(* IEC 61131-3 sources: daoli-st-library/DL_Base (part 15) *)

(* ---- FB_DL_RailPowerSequence.st ---- *)
(*
  ==================================================================
  组件名 Component  : FB_DL_RailPowerSequence
  分类   Category   : DL_Base
  前缀   Naming     : FB_DL_ ｜ b/n/u/f/t/e/st 类型前缀制（R265）
  复杂度 Complexity  : 中
  版本   Version    : 1.0.3
  功能   Purpose    : 多路供电轨按序上电/断电（延时可配、断电逆序、步进超时锁存）。
  来源   Source     : self-std（供电时序公开工程语义自研）
  平台   Platform   : 纯 IEC 61131-3（TON / R_TRIG / CASE），三平台通用
  分工声明 Split     : 与 FB_DL_LaserWeldPowerSeq（工艺专用属主）分工——后者绑定
                      激光焊接工艺流；本件为通用时序原子，不绑工艺、不判负载
                      特性（R216 双向互引）。
  作者   Author     : 道莅代码库 · PLC 编程专家（R61）
  归属 Ownership     : E_DL_RailPhase 属主为本文件（全库唯一定义，R264）；
                      引用件只引用不重声明。
  ------------------------------------------------------------------
  边界 Boundary     :
                      一 uRailCount = 0 或 > 8 判组态非法故障码，不进时序
                         （边界五；R239 显式分支，禁比较算子隐式分流）；
                      二 断电逆序强制：断电步序 = 上电步序倒序（结构写死）；
                      三 步进超时按「单轨」计时（v1.0.2 修 D2）：tonStep.IN 串入逐拍派生
                         的本轨待响应量 _bRailPending（eRampUp 取 NOT abRailFb[_nStep]、
                         eRampDn 取 abRailFb[_nStep]），本轨一响应即自动复位，不再整段
                         连续计时；锁存独立码 + 解除式可达自证：故障相由复位沿迁回空闲
                         并清锁存（bReset 输入引脚恒可达，R152 自证）；
                      三A 上电推进判据「沿 OR 电平」双路（v1.0.3 修 R62-D4 中）：eRampUp
                         推进条件 = rtFb.Q（反馈上升沿）OR abRailFb[_nStep]（电平已就位
                         直过）——「反馈预闭合」处置口径：若轨在上一步计时期间或起步拍
                         前反馈电平已提前闭合（边沿被上一步消费 / 起步拍无沿），单轨超时
                         门控（_bRailPending = FALSE）与推进判据（仅沿）同源失效会静默
                         挂死；电平直过支路消除该挂死路径。断电相完成判据本为电平式
                         （NOT abRailFb[_nStep]），无此问题；
                      七 空轨断电早退（v1.0.2 修 D1）：_nCnt = 0 时收到断电沿不迁移、
                         不置 bDone、仅发信息级 0655，防伪造「完成单拍」；原负下标
                         钳位语句保留为二重防御，不再是唯一防线；
                      四 状态机 ENUM + CASE，ELSE 拦非法态；TON/R_TRIG 段 0
                         无条件刷新（禁入分支，R7）；TON IN 串故障锁存门控
                         （FB50-1）；
                      五 使能失电语义为「弃用本轮时序」（回空闲，不锁存不出
                         单拍）——R191 声明行；
                      六 无全局、无外部变量、无物理地址。
  错误码   Codes    :
    16#0001_0642【故障级】供电轨数组态非法（=0 或 >8），锁存至复位沿
    16#0001_0643【故障级】步进反馈超时（tStepTimeout 内未见该轨反馈），锁存至复位沿
    16#0001_0655【信息级】空轨断电请求已忽略（_nCnt 为 0 时无可断轨，不迁移不置 bDone）
  验收   Acceptance :
    算法已证（脚本）：未跑 ｜ 编译器已证（三平台）：未跑
    V1 3 轨、反馈逐轨到位 → uOnCount=3、bDone 单拍
    V2 第 2 轨反馈不至 → 码 0643、eFault、锁存待复位
    V3 uRailCount=0 → 码 0642、不进时序
    V4 空轨断电（abRailFb 全 FALSE、bOffCmd 上升沿）→ bDone 全拍 FALSE、
       eState 保持 eIdle、eErr=0655（v1.0.2 回归向量）
    V5 3 轨、每轨反馈延时 0.8×tStepTimeout → 全序列成功、无 0643；
       单轨延时 1.2× → 该轨锁 0643（v1.0.2 单轨超时回归向量）
    V6 轨 2 反馈预闭合（在轨 1 计时期间电平提前拉高，无沿）→ 轨 2 仍被推进、
       不锁 0643（v1.0.3 沿 OR 电平双路回归向量）
  修订记录 Revision  :
    2026-11-21  v1.0.0  R61 首版（批 3 · 序号 9）
    2026-11-21  v1.0.1  R61 终审 D1 就地修（安全侧）：空轨断电起步 _nStep<0 钳位、堵 abRailFb[-1] 越界读（R333 安全侧例外，正常路径行为零变更）
    2026-11-21  v1.0.2  R62-D1/D2 返修：①eIdle/eStable 的 rtOff 分支加 _nCnt=0 空轨早退（不迁移、不置 bDone、仅信息码 0655），原钳位降为二重防御；②新增 _bRailPending 串入 tonStep.IN 实现单轨超时；③段 0 rtFb 刷新条件扩到 eRampUp 或 eRampDn
    2026-11-21  v1.0.3  R63 返修 R4（R62-D4 中）：eRampUp 推进判据改「沿 OR 电平」双路（rtFb.Q OR abRailFb[_nStep]），反馈预闭合轨电平直过，消除单轨超时门控与推进判据同源静默挂死；头注释补「反馈预闭合」处置口径与向量 V6
  ==================================================================
*)
TYPE E_DL_RailPhase :
(
    eIdle    := 0,  // 空闲：等上电/断电命令沿 / idle, waiting for the power command edges
    eRampUp  := 10, // 上电步进：正向逐轨 / the power up stepping forward rail by rail
    eStable  := 20, // 稳定：全轨已上 / stable, all rails powered
    eRampDn  := 30  // 断电步进：逆向逐轨（边界二）/ the power down stepping in the reverse order
);
END_TYPE

FUNCTION_BLOCK FB_DL_RailPowerSequence
VAR_INPUT
    bOnCmd       : BOOL := FALSE; // 上电命令电平，上升沿发起正向时序 / the power on command level
    bOffCmd      : BOOL := FALSE; // 断电命令电平，上升沿发起逆向时序 / the power off command level
    bReset       : BOOL := FALSE; // 故障复位电平，上升沿清锁存回空闲 / the fault reset level
    uRailCount   : UDINT := 3;    // 供电轨数 [路]，合法域 1..8 / the rail count, legal from one to eight
    tStepTimeout : TIME := T#5S;  // 单轨步进超时 [毫秒] / the per rail step timeout
END_VAR
VAR_IN_OUT
    abRailFb  : ARRAY[0..7] OF BOOL; // 各轨反馈电平 [路反馈]，只读 / the rail feedback levels, read only
    atOnDelay : ARRAY[0..7] OF TIME; // 各轨上电前延时 [毫秒]，可配 / the per rail pre power delay, configurable
END_VAR
VAR_OUTPUT
    uOnCnt  : UDINT := 0;              // 已上电轨数 [路] / the powered rail count
    bDone   : BOOL := FALSE;           // 本轮时序完成单拍脉冲 [-] / the round done one shot pulse
    eState  : E_DL_RailPhase;          // 主状态机当前态 [状态] / the current state
    bError  : BOOL := FALSE;           // 故障锁存位（与锁存同源，R191）/ the fault bit from the latch
    eErr    : UDINT := 16#0000_0000;   // 错误码，0 = 正常 / the error code, zero is ok
END_VAR
VAR
    _bInit   : BOOL := FALSE;                          // 首拍初始化标志（R310）/ the first scan flag
    _eState  : E_DL_RailPhase := E_DL_RailPhase.eIdle; // 内部状态寄存器 / the internal state register
    _bDone   : BOOL := FALSE;                          // 完成单拍内部位，段 1 预清段 5 映射 / the internal done bit
    _bFault  : BOOL := FALSE;                          // 故障锁存副本（仅复位沿清除）/ the fault latch copy
    _nStep   : DINT  := 0;                             // 当前步进轨索引 [下标] / the current step rail index
    _nCnt    : UDINT := 0;                             // 已完成轨数副本 [路] / the completed rail count copy
    _nUse    : DINT  := 0;                             // 钳位后的轨数 [路] / the clamped rail count
    _bCfgBad : BOOL  := FALSE;                         // 组态非法标记（逐拍重算）/ the configuration fault flag
    _bStepGo : BOOL  := FALSE;                         // 步进计时使能（驻留派生）[-] / the step timing enable derived from the dwell
    _bRailPending : BOOL := FALSE;                     // 本轨待响应量（逐拍派生：上电取未反馈、断电取仍反馈）[-] / the pending rail of this step, derived every scan
    _bEmptyOff : BOOL := FALSE;                        // 空轨断电早退标记（逐拍重算，信息级 0655）/ the empty bank off request flag, recomputed every scan
    rtOn     : R_TRIG;  // 上电命令沿实例，段 0 无条件刷新 / the on command edge instance
    rtOff    : R_TRIG;  // 断电命令沿实例，段 0 无条件刷新 / the off command edge instance
    rtReset  : R_TRIG;  // 复位沿实例，段 0 无条件刷新 / the reset edge instance
    rtFb     : R_TRIG;  // 步进轨反馈沿实例，段 0 无条件刷新 / the step rail feedback edge instance
    tonStep  : TON;     // 步进超时计时器，段 0 无条件刷新 / the step timeout timer
END_VAR
VAR CONSTANT
    DL_RPS_RMAX : DINT := 8; // 供电轨容量上界 [路]，与数组容量一致 / the rail capacity aligned with the array
END_VAR

// 段 0｜定时器与沿检测无条件周期刷新（禁入分支，R7；TON IN 串故障锁存门控，FB50-1）/ segment 0, the unconditional refresh
rtOn(CLK := bOnCmd); // 上电沿 / the on edge
rtOff(CLK := bOffCmd); // 断电沿 / the off edge
rtReset(CLK := bReset); // 复位沿 / the reset edge
IF (_eState = E_DL_RailPhase.eRampUp) OR (_eState = E_DL_RailPhase.eRampDn) THEN // 两相步进相均刷当前轨反馈（v1.0.2 扩相，防断电相恒刷 0 号轨）/ both stepping phases watch the current rail
    rtFb(CLK := abRailFb[_nStep]); // 当前步进轨反馈沿 / the current step rail feedback edge
ELSE // 非步进相：非步进相固定刷新 0 号轨（保持无条件调用形态）/ the other phases refresh on the rail zero slot
    rtFb(CLK := abRailFb[0]); // 固定下标刷新 / the fixed index refresh
END_IF
_bStepGo := (_eState = E_DL_RailPhase.eRampUp) OR (_eState = E_DL_RailPhase.eRampDn); // 步进相驻留派生 / the dwell derived enable
// 单轨待响应量：只由「本相 + 本轨反馈」派生，本轨一响应即落 FALSE 使 TON 自动复位（v1.0.2 修 D2）/ the per rail pending, the timer resets by itself once this rail responds
IF _eState = E_DL_RailPhase.eRampUp THEN // 上电相：本轨尚未反馈即待响应 / the ramp up phase waits for the feedback to appear
    _bRailPending := NOT abRailFb[_nStep]; // 未反馈为待响应 / pending while the feedback is still absent
ELSIF _eState = E_DL_RailPhase.eRampDn THEN // 断电相：本轨仍反馈即待响应 / the ramp down phase waits for the feedback to vanish
    _bRailPending := abRailFb[_nStep]; // 仍反馈为待响应 / pending while the feedback is still present
ELSE // 其余相无单轨待响应语义 / no per rail pending outside the stepping phases
    _bRailPending := FALSE; // 非步进相清待响应 / clear the pending outside the stepping phases
END_IF
tonStep(IN := _bStepGo AND (NOT _bFault) AND _bRailPending, PT := tStepTimeout); // 单轨超时（串故障锁存门控 + 本轨待响应，FB50-1）/ the per rail timeout with the latch gate and the rail pending

// 段 1｜首拍初始化与单拍标志预清（FB32-1；R256）/ segment 1, the first scan init and the preset
IF NOT _bInit THEN // 首拍一拍 / the first scan
    _bInit := TRUE; // 置首拍标志 / raise the first scan flag
    _bFault := FALSE; // 故障锁存显式清零 / clear the fault latch explicitly
    _nStep := 0; // 步进索引显式清零 / clear the step index explicitly
    _nCnt := 0; // 完成轨数显式清零 / clear the completed count explicitly
    _eState := E_DL_RailPhase.eIdle; // 状态显式落空闲 / place the state to idle
END_IF
IF rtReset.Q THEN // 复位沿（作用域：清锁存 + 迁相位 + 清步进量，R311）/ the reset edge with the declared scope
    _bFault := FALSE; // 清故障锁存 / clear the fault latch
    _nStep := 0; // 清步进索引 / clear the step index
    _nCnt := 0; // 清完成轨数 / clear the completed count
    _eState := E_DL_RailPhase.eIdle; // 迁回空闲 / back to idle
END_IF
_bDone := FALSE; // 完成单拍预清零 / preset the done pulse false
_bCfgBad := FALSE; // 组态标记预清零 / preset the configuration flag false
_bEmptyOff := FALSE; // 空轨早退标记预清零（单拍信息位，段 5 映射 0655）/ preset the empty bank flag false

// 段 2｜组态域闸（轨数合法域 1..8，边界一）/ segment 2, the rail count gate
_nUse := UDINT_TO_DINT(uRailCount); // 轨数升位接管（超 DINT 域转负即被下界捕获）/ take the rail count widened, an overflow lands below the floor
IF (_nUse < 1) OR (_nUse > DL_RPS_RMAX) THEN // 轨数越域 / the rail count out of the domain
    _bCfgBad := TRUE; // 置组态非法标记 / raise the configuration flag
    _bFault := TRUE; // 锁存故障（0642，段 5 回放）/ latch the fault
END_IF
IF _nUse < 1 THEN // 下界钳位（防越界索引）/ the floor clamp for the index safety
    _nUse := 1; // 钳到一 / clamp to one
END_IF
IF _nUse > DL_RPS_RMAX THEN // 上界钳位 / the ceiling clamp
    _nUse := DL_RPS_RMAX; // 钳到容量 / clamp to the capacity
END_IF

// 段 3｜主状态机（ENUM + CASE，ELSE 拦非法态；安全相迁移带全量闸位复检，R274）/ segment 3, the main machine
CASE _eState OF
    E_DL_RailPhase.eIdle: // 空闲相 / the idle phase
        IF rtOn.Q AND (NOT _bFault) AND (NOT _bCfgBad) THEN // 上电沿 + 全量闸位复检（R274）/ the on edge with the full gate recheck
            _nStep := 0; // 从 0 号轨正向起步 / start forward from the rail zero
            _nCnt := 0; // 完成轨数归零 / reset the completed count
            _eState := E_DL_RailPhase.eRampUp; // 迁入上电步进相 / enter the ramp up phase
        ELSIF rtOff.Q AND (NOT _bFault) AND (NOT _bCfgBad) THEN // 断电沿 + 全量闸位复检 / the off edge with the recheck
            IF _nCnt = 0 THEN // 空轨早退（v1.0.2 修 D1）：无已上电轨则无从逆序断电 / the empty bank early exit, no powered rail to cut
                _bEmptyOff := TRUE; // 仅置信息级标记，不迁移、不置 bDone / raise the informational flag only, no migration and no done pulse
            ELSE // 有已上电轨：正常逆序起步 / a powered bank, start the reverse sequence
                _nStep := UDINT_TO_DINT(_nCnt) - 1; // 从已完成末轨逆向起步（断电逆序，边界二）/ start reverse from the last powered rail
                IF _nStep < 0 THEN // 二重防御：空轨已在上面早退，本钳位不再是唯一防线（R61-D1 保留）/ a second line of defence, no longer the only guard
                    _nStep := 0; // 钳到 0 号轨，防 abRailFb[-1] 越界读 / clamp to the rail zero against the negative index read
                END_IF
                _eState := E_DL_RailPhase.eRampDn; // 迁入断电步进相 / enter the ramp down phase
            END_IF
        END_IF
    E_DL_RailPhase.eRampUp: // 上电步进相 / the ramp up phase
        IF rtFb.Q OR abRailFb[_nStep] THEN // 推进判据「沿 OR 电平」双路（v1.0.3 修 R62-D4）：沿到或电平已预闭合均直过，防超时门控与推进判据同源静默挂死 / the advance criterion in the edge OR level dual path, a pre closed feedback passes by level so the timeout gate and the advance criterion cannot fail together in silence
            _nCnt := _nCnt + 1; // 完成轨数推进 / advance the completed count
            _nStep := _nStep + 1; // 步进索引推进 / advance the step index
            IF _nStep >= _nUse THEN // 全轨完成 / all rails done
                _bDone := TRUE; // 置完成单拍 / raise the done pulse
                _eState := E_DL_RailPhase.eStable; // 迁入稳定相 / enter the stable phase
            END_IF
        ELSIF tonStep.Q THEN // 步进超时（边界三）/ the step timeout
            _bFault := TRUE; // 锁存超时故障（0643）/ latch the timeout fault
        ELSIF _bFault THEN // 前置条件消失出口 / the prerequisite gone exit
            _eState := E_DL_RailPhase.eIdle; // 迁回空闲（锁存迁移由段 4 收口）/ back to idle
        END_IF
    E_DL_RailPhase.eStable: // 稳定相 / the stable phase
        IF rtOff.Q AND (NOT _bFault) THEN // 断电沿 + 闸位复检 / the off edge with the recheck
            IF _nCnt = 0 THEN // 空轨早退（与 eIdle 同口径，v1.0.2 修 D1）：异常态下 _nCnt 被清零亦不得伪造完成 / the same empty bank exit as the idle phase
                _bEmptyOff := TRUE; // 仅置信息级标记，不迁移、不置 bDone / raise the informational flag only
            ELSE // 有已上电轨：正常逆序起步 / a powered bank, start the reverse sequence
                _nStep := UDINT_TO_DINT(_nCnt) - 1; // 逆向起步（断电逆序）/ start reverse
                IF _nStep < 0 THEN // 二重防御（空轨已在上面早退）/ a second line of defence
                    _nStep := 0; // 钳到 0 号轨，防负下标越界读 / clamp to the rail zero against the negative index read
                END_IF
                _eState := E_DL_RailPhase.eRampDn; // 迁入断电步进相 / enter the ramp down phase
            END_IF
        ELSIF _bFault THEN // 前置条件消失 / the prerequisite gone
            _eState := E_DL_RailPhase.eIdle; // 迁回空闲 / back to idle
        END_IF
    E_DL_RailPhase.eRampDn: // 断电步进相（逆序，边界二）/ the ramp down phase in the reverse order
        IF NOT abRailFb[_nStep] THEN // 当前轨反馈已消失（断电完成判据）/ the current rail feedback gone
            IF _nCnt > 0 THEN // 无符号下溢闸（0 减 1 会回绕，先判再减）/ the underflow guard before the decrement
                _nCnt := _nCnt - 1; // 完成轨数回退 / step the completed count back
            END_IF
            _nStep := _nStep - 1; // 逆向推进 / step reverse
            IF _nStep < 0 THEN // 全轨断完 / all rails off
                _nCnt := 0; // 完成轨数清零 / clear the completed count
                _bDone := TRUE; // 置完成单拍 / raise the done pulse
                _eState := E_DL_RailPhase.eIdle; // 迁回空闲 / back to idle
            END_IF
        ELSIF tonStep.Q THEN // 步进超时 / the step timeout
            _bFault := TRUE; // 锁存超时故障 / latch the timeout fault
        ELSIF _bFault THEN // 前置条件消失 / the prerequisite gone
            _eState := E_DL_RailPhase.eIdle; // 迁回空闲 / back to idle
        END_IF
    ELSE // 非法枚举值拦截 / the illegal enumeration guard
        _eState := E_DL_RailPhase.eIdle; // 落回空闲 / force back to idle
        _bFault := TRUE; // 置故障锁存 / latch the fault
END_CASE

// 段 4｜故障锁存迁移闸（置于解除段之后防同拍抢迁，R258）/ segment 4, the latch to phase gate
IF _bFault AND (_eState <> E_DL_RailPhase.eIdle) THEN // 已锁存但不在空闲相（本件锁存即弃用本轮迁空闲）/ latched, the round is discarded to idle
    _eState := E_DL_RailPhase.eIdle; // 迁回空闲 / back to idle
END_IF

// 段 5｜统一出口（内部副本单点映射；故障码锁存回放，R187）/ segment 5, the unified outlet
uOnCnt := _nCnt; // 已上电轨数出口 / the powered count outlet
bDone := _bDone; // 完成单拍出口 / the done pulse outlet
eState := _eState; // 状态出口 / the state outlet
bError := _bFault; // 故障位出口（与锁存同源）/ the fault bit outlet
IF _bFault THEN // 故障锁存回放优先 / the latched fault replays first
    IF _bCfgBad THEN // 组态成因（独立码值，R190）/ the configuration cause
        eErr := 16#0001_0642; // 故障级：轨数组态非法 / fault grade, the illegal rail count
    ELSE // 超时成因 / the timeout cause
        eErr := 16#0001_0643; // 故障级：步进反馈超时 / fault grade, the step feedback timeout
    END_IF
ELSE // 无故障 / no fault
    IF _bEmptyOff THEN // 空轨断电请求已忽略（信息级不置 bError，R285）/ the empty bank request ignored, informational without bError
        eErr := 16#0001_0655; // 信息级：空轨断电请求已忽略 / informational, the empty bank off request ignored
    ELSE // 无事件 / no event
        eErr := 16#0000_0000; // 正常 / ok
    END_IF
END_IF
END_FUNCTION_BLOCK

(* ---- FB_DL_RecipeStepExec.st ---- *)
(*
    FB_DL_RecipeStepExec —— 配方步序执行器（步推进 / 步超时 / 暂停恢复 / 禁跳步）
    ------------------------------------------------------------------
    组件名称  : FB_DL_RecipeStepExec
    分类      : DL_Base / Sequencing
    前缀      : FB_DL_
    版本      : 1.0.0
    溯源      : 借鉴点 —— PackML / ISA-TR88.00.02 状态模型的「执行态 + 保持（暂停）态 +
                完成态 + 中止」四类状态语义，以及配方步序「逐步等待动作完成信号」
                的通行做法；步超时、暂停恢复、禁跳步三项为工程惯例约束。
                本件只借鉴**状态语义与约束项**，不借用其状态表实现。
                clean-room 声明 —— 零代码行复制；状态机为本件自有 ENUM + CASE，
                定时仅用 IEC 61131-3 标准库 TON，沿检测仅用标准库 R_TRIG。
                许可证 —— 本件 MIT；来源标签 packml 指标准状态模型术语，
                标准文本不属代码，无许可继承。
    平台      : 纯 IEC 61131-3，CODESYS 3.5 / TwinCAT 3 / InoProShop / Machine Expert 通用
    作者      : 道莅代码库 · PLC编程专家（R70 构建轮 · 批 3 · N9）
    ------------------------------------------------------------------
    功能说明  : 步号从 1 走到 nStepTotal。每步等待 bStepDone 上升沿推进，
                推进即「步号 + 1」；超过 nStepTotal 则完成。
                步超时：_tonStep 的 PT = tStep，IN = 运行态 且 非「步切换复位拍」；
                步号一旦切换（推进 / 跳步 / 暂停恢复）就置 _bTimerRestart，
                使下一拍 IN 断开一拍、计时器复位、本步重新从 0 计时 —— 若不这样做，
                计时器会跨步累计，第二步必然立刻超时（历史教训：定时器不自复位）。
                暂停恢复：bPause 为电平（TRUE 即暂停）。暂停期间步超时计时**复位**
                （IN 断开），恢复后本步重新计时；该语义写死于边界三，不留歧义。
                禁跳步：仅允许跳到「当前步 + 1」（等价于立即完成本步）；其余目标
                一律拒绝，置信息级码 0703，bError 保持 FALSE，状态与步号不变。
    错误码    : 16#0002_0701 组态非法（nStepTotal < 1 或 tStep <= T#0S），锁存 —— 故障级
                16#0002_0702 步超时（当前步未在 tStep 内收到完成信号），锁存 —— 故障级
                16#0002_0703 跳步被拒（目标非「当前步 + 1」或越出总量），不锁存 —— 信息级
                16#0002_0704 非法状态枚举值（CASE ELSE 兜底），锁存 —— 故障级
    码位总账  : 0701 / 0702 / 0704 用（故障级，锁存回放）｜ 0703 用（信息级，每拍重算）
    状态机    : ENUM E_DL_RseState 五态，CASE 全覆盖 + ELSE 兜底（回 eFault 置 0704）。
                迁移：eIdle -启动沿-> eRun -完成-> 步号+1（超总量 -> eDone）
                      eRun -bPause-> ePause -NOT bPause-> eRun
                      任意态 -bAbort-> eIdle（操作态，不发码）
                      任意态 -锁存故障-> eFault；eFault -bReset 沿-> eIdle（唯一解除边）
    边界与披露: 一 组态闸（R272 逐项点名）：nStepTotal < 1 拦截（无步可执行）；
                   tStep <= T#0S 拦截（零超时使第一步即失败，属组态错误）；
                二 输入闸：nJumpTo 为整型无 NaN 面，按 1..nStepTotal 区间校验，
                   越界即判为「跳步被拒」，不参与任何数组索引（本件无数组）；
                三 暂停恢复语义（R191 声明）：暂停期间步超时计时器复位，恢复后
                   本步从头计时 —— 即「暂停不计入步超时」，这是本件的判定口径；
                四 失能语义：本件无 bEn 引脚，停机由 bAbort 承担（电平有效），
                   bAbort 为真即回 eIdle 且步号清零、bStepActive / bPaused / bDone
                   全清零，不发码（操作态）；
                五 单拍位口径（R256）：bJumpRejected 为单拍信息位，段 1 统一预置，
                   仅在被拒的那一拍由 CASE 置真；bDone 为保持位（完成态持续为真）；
                六 定时器 _tonStep 与四个沿实例 _rtStart / _rtReset / _rtDone / _rtJump
                   全部每周期无条件调用（规则 ⑦）；
                七 零全局变量、零 VAR_EXTERNAL、零物理地址、零除法、零数组下标。
    修订记录  : 2026-11-22 v1.0.0 首次入库（R70 构建轮 · 批 3 · N9）
*)
TYPE E_DL_RseState :
(
    eIdle  := 0,   (* 待机，等待启动 / idle, waiting for a start *)
    eRun   := 10,  (* 执行态（某一步激活中）/ running, a step is active *)
    ePause := 20,  (* 暂停态（步保持，超时计时复位）/ paused, the step holds and its timer resets *)
    eDone  := 30,  (* 完成态（全部步执行完毕，保持）/ done, every step finished, held *)
    eFault := 40   (* 故障态（锁存待复位）/ fault, latched for a reset *)
);
END_TYPE

FUNCTION_BLOCK FB_DL_RecipeStepExec
VAR_INPUT
    bStart     : BOOL := FALSE;            (* 启动序列（上升沿有效），[标志] / the sequence start, rising edge *)
    bStepDone  : BOOL := FALSE;            (* 当前步动作完成（上升沿有效），[标志] / the current step finished, rising edge *)
    bPause     : BOOL := FALSE;            (* 暂停（电平有效，TRUE 即暂停），[标志] / the pause, level effective *)
    bAbort     : BOOL := FALSE;            (* 中止（电平有效），[标志] / the abort, level effective *)
    bReset     : BOOL := FALSE;            (* 故障复位（上升沿有效），[标志] / the fault reset, rising edge *)
    bJumpReq   : BOOL := FALSE;            (* 跳步请求（上升沿有效），[标志] / the jump request, rising edge *)
    nJumpTo    : INT := 0;                 (* 跳步目标步号，[号]，域 1..nStepTotal / the jump target step number *)
    nStepTotal : INT := 10;               (* 步总数，[步]，须 >= 1 / the total number of steps, must be at least one *)
    tStep      : TIME := T#30S;            (* 单步超时，[ms]，须 > T#0S / the per step timeout *)
END_VAR
VAR_OUTPUT
    eState      : E_DL_RseState := E_DL_RseState.eIdle; (* 状态出口，[状态] / the state outlet *)
    nStepNo     : INT;                     (* 当前步号，0 = 无步激活，[号] / the current step number, 0 = none *)
    bStepActive : BOOL;                    (* 当前步激活中，[标志] / the current step is active *)
    bPaused     : BOOL;                    (* 暂停中，[标志] / paused *)
    bDone       : BOOL;                    (* 序列完成（保持），[标志] / the sequence completed, held *)
    bJumpRejected : BOOL;                  (* 跳步被拒单拍位，[标志] / the jump was rejected, single scan *)
    bBusy       : BOOL;                    (* 序列占用中（执行或暂停），[标志] / the sequence is occupied *)
    bValid      : BOOL;                    (* 出口可信（非故障态），[标志] / the outlets are trustworthy *)
    bError      : BOOL;                    (* 故障标志，故障级码时为 TRUE / the error flag, TRUE on fault level *)
    nErrCode    : UDINT;                   (* 错误码，0 = 正常 / the error id, 0 = ok *)
END_VAR
VAR
    _rtStart     : R_TRIG;                 (* 启动上升沿实例（无条件调用）/ the start edge instance *)
    _rtReset     : R_TRIG;                 (* 复位上升沿实例（无条件调用）/ the reset edge instance *)
    _rtDone      : R_TRIG;                 (* 步完成上升沿实例（无条件调用）/ the step done edge instance *)
    _rtJump      : R_TRIG;                 (* 跳步请求上升沿实例（无条件调用）/ the jump request edge instance *)
    _tonStep     : TON;                    (* 步超时计时实例（无条件调用）/ the step timeout timer *)
    _eState      : E_DL_RseState := E_DL_RseState.eIdle; (* 状态寄存器，[状态] / the internal state register *)
    _nStep       : INT;                    (* 当前步号寄存器，[号] / the internal step register *)
    _bFault      : BOOL;                   (* 故障锁存位，仅 bReset 上升沿解除 / the latched fault bit *)
    _nCodeLatch  : UDINT;                  (* 锁存成因码，故障期回放 / the latched cause code *)
    _bCfgBad     : BOOL;                   (* 组态非法标志（逐拍重算）/ the configuration fault flag *)
    _bTimerIn    : BOOL;                   (* 步计时器 IN 条件（显式条件）/ the timer IN condition *)
    _bTimerRestart : BOOL;                 (* 步切换复位拍标志（使计时器下一拍复位）/ the timer restart flag *)
    _bJumpOk     : BOOL;                   (* 跳步目标合法标志，[标志] / the jump target is legal *)
    _bAdvanced   : BOOL;                   (* 本拍发生过步号推进，[标志] / the step advanced this scan *)
END_VAR

// 段 1｜出口预置（R256 统一出口预置，单拍位在此清零）/ segment 1, preset every outlet
eState       := _eState;                   // 状态出口先镜像寄存器 / mirror the state register first
nStepNo      := _nStep;                    // 步号出口先镜像寄存器 / mirror the step register first
bStepActive  := FALSE;                     // 步激活位预清零 / preset the step active flag false
bPaused      := FALSE;                     // 暂停位预清零 / preset the paused flag false
bDone        := FALSE;                     // 完成位预清零（保持态另由 eDone 分支置真）/ preset the done flag false
bJumpRejected := FALSE;                    // 跳步被拒单拍位预清零（R256）/ preset the jump rejected flag false
bBusy        := FALSE;                     // 占用标志预清零 / preset the busy flag false
bValid       := TRUE;                      // 可用标志预置真（故障态再清）/ preset valid true
bError       := FALSE;                     // 故障标志预清零 / preset the error flag false
nErrCode     := 0;                         // 错误码预置无错 / preset the code to zero
_bAdvanced   := FALSE;                     // 推进标志预清零 / preset the advanced flag false

// 段 2｜沿实例与定时器无条件周期调用（规则 ⑦）/ segment 2, the edges and the timer, called unconditionally
_rtStart(CLK := bStart);                   // 启动沿，每周期无条件刷新 / the start edge, refreshed every scan
_rtReset(CLK := bReset);                   // 复位沿，每周期无条件刷新 / the reset edge, refreshed every scan
_rtDone(CLK := bStepDone);                 // 步完成沿，每周期无条件刷新 / the step done edge, refreshed every scan
_rtJump(CLK := bJumpReq);                  // 跳步沿，每周期无条件刷新 / the jump edge, refreshed every scan
_bTimerIn := (_eState = E_DL_RseState.eRun) AND NOT _bTimerRestart; // 运行态且非复位拍才计时
_tonStep(IN := _bTimerIn, PT := tStep);    // 步超时计时，每周期无条件调用 / the step timeout timer
_bTimerRestart := FALSE;                   // 复位拍已消费，本拍清标志 / the restart flag is consumed

// 段 3｜复位解除：唯一可到达的清除边（R188）/ segment 3, the only latch release edge
IF _rtReset.Q THEN                         // 复位上升沿 / the reset rising edge
    _bFault     := FALSE;                  // 解除故障锁存 / release the fault latch
    _nCodeLatch := 0;                      // 清锁存码 / clear the latched code
    _eState     := E_DL_RseState.eIdle;    // 回待机（安全相）/ back to the safe idle phase
    _nStep      := 0;                      // 步号清零 / clear the step number
    _bTimerRestart := TRUE;                // 计时器下一拍复位 / restart the timer next scan
END_IF

// 段 4｜组态守卫（R272 逐项点名）/ segment 4, the configuration guard
_bCfgBad := (nStepTotal < 1) OR (tStep <= T#0S); // 步总数为零 或 超时非正 / no steps or a non positive timeout

// 段 5｜首次成因锁存（故障期不重推断，R189）/ segment 5, the first cause latch
IF NOT _bFault THEN                        // 未锁存才登记 / register only while healthy
    IF _bCfgBad THEN                       // 组态非法 / an illegal configuration
        _bFault     := TRUE;               // 置锁存 / latch it
        _nCodeLatch := 16#0002_0701;       // 故障级：组态非法 / fault level: an illegal configuration
        _eState     := E_DL_RseState.eFault; // 迁入故障态 / enter the fault state
    END_IF
END_IF

// 段 6｜中止命令（操作态，不发码）/ segment 6, the abort command
IF bAbort AND NOT _bFault THEN             // 中止有效且无锁存故障 / an abort without a latched fault
    _eState := E_DL_RseState.eIdle;        // 回待机 / back to idle
    _nStep  := 0;                          // 步号清零 / clear the step number
END_IF

// 段 7｜状态机（ENUM + CASE + ELSE 兜底）/ segment 7, the state machine
CASE _eState OF
    E_DL_RseState.eIdle:                   // 待机态 / the idle state
        bValid := TRUE;                    // 待机出口可信 / the idle outlets are trustworthy
        IF _rtStart.Q AND NOT _bFault THEN // 启动沿且无锁存故障 / a start edge without a latched fault
            _nStep  := 1;                  // 从第 1 步开始 / start from step one
            _eState := E_DL_RseState.eRun; // 进入执行态 / enter the running state
            _bTimerRestart := TRUE;        // 计时器下一拍复位（本步从 0 计时）/ restart the timer for the new step
        END_IF
    E_DL_RseState.eRun:                    // 执行态 / the running state
        bStepActive := TRUE;               // 当前步激活 / the step is active
        bBusy       := TRUE;               // 序列占用 / the sequence is occupied
        IF bPause THEN                     // 暂停命令（电平）/ the pause command, level
            _eState := E_DL_RseState.ePause; // 进入暂停态 / enter the paused state
        ELSIF _rtJump.Q THEN               // 跳步请求沿 / a jump request edge
            IF (nJumpTo >= 1) AND (nJumpTo <= nStepTotal) AND (nJumpTo = (_nStep + 1)) THEN
                _bJumpOk := TRUE;          // 目标为「当前步 + 1」，合法 / the target is the next step, legal
            ELSE                           // 其余目标一律拒绝（禁跳步）/ every other target is refused
                _bJumpOk := FALSE;         // 非法目标 / an illegal target
            END_IF
            IF _bJumpOk THEN               // 合法跳步 / a legal jump
                IF _nStep >= nStepTotal THEN // 已是最后一步 / already the last step
                    _eState := E_DL_RseState.eDone; // 进入完成态 / enter the done state
                ELSE                       // 非最后一步 / not the last step
                    _nStep := _nStep + 1;  // 步号推进 / advance the step
                    _bAdvanced := TRUE;    // 标记推进 / mark the advance
                END_IF
            ELSE                           // 跳步被拒 / the jump is refused
                bJumpRejected := TRUE;     // 单拍被拒位（R256）/ the single scan rejected flag
                nErrCode      := 16#0002_0703; // 信息级：跳步被拒（不置 bError，R45）/ info level, no fault flag
            END_IF
        ELSIF _rtDone.Q THEN               // 步完成沿 / the step done edge
            IF _nStep >= nStepTotal THEN   // 最后一步完成 / the last step finished
                _eState := E_DL_RseState.eDone; // 进入完成态 / enter the done state
            ELSE                           // 非最后一步 / not the last step
                _nStep := _nStep + 1;      // 步号推进 / advance the step
                _bAdvanced := TRUE;        // 标记推进 / mark the advance
            END_IF
        ELSIF _tonStep.Q THEN              // 步超时 / the step timed out
            _bFault     := TRUE;           // 锁存故障 / latch the fault
            _nCodeLatch := 16#0002_0702;   // 故障级：步超时 / fault level: a step timeout
            _eState     := E_DL_RseState.eFault; // 迁入故障态 / enter the fault state
        END_IF
    E_DL_RseState.ePause:                  // 暂停态 / the paused state
        bStepActive := TRUE;               // 步保持（不推进也不超时）/ the step holds, neither advanced nor timed
        bPaused     := TRUE;               // 暂停标志 / the paused flag
        bBusy       := TRUE;               // 序列仍占用 / the sequence is still occupied
        IF NOT bPause THEN                 // 暂停解除 / the pause released
            _eState := E_DL_RseState.eRun; // 回执行态 / back to running
            _bTimerRestart := TRUE;        // 本步重新计时（边界三口径）/ the step is timed from zero again
        END_IF
    E_DL_RseState.eDone:                   // 完成态（保持）/ the done state, held
        bDone  := TRUE;                    // 完成标志 / the done flag
        bValid := TRUE;                    // 完成态出口可信 / the done outlets are trustworthy
        IF _rtStart.Q THEN                 // 再次启动 = 新一轮 / a new start begins a new run
            _nStep  := 1;                  // 回到第 1 步 / back to step one
            _eState := E_DL_RseState.eRun; // 进入执行态 / enter the running state
            _bTimerRestart := TRUE;        // 计时器复位 / restart the timer
        END_IF
    E_DL_RseState.eFault:                  // 故障态（锁存保持）/ the fault state, latched
        bValid   := FALSE;                 // 出口不可信 / the outlets are not trustworthy
        bError   := TRUE;                  // 故障标志置位 / raise the fault flag
        nErrCode := _nCodeLatch;           // 回放锁存码 / replay the latched code
    ELSE                                   // 非法枚举兜底（回安全相 + 置码，规则 ⑥）/ the illegal enumeration guard
        _bFault     := TRUE;               // 置锁存 / latch it
        _nCodeLatch := 16#0002_0704;       // 故障级：非法状态枚举 / fault level: an illegal state value
        _eState     := E_DL_RseState.eFault; // 回安全相 / force the safe fault state
        bValid      := FALSE;              // 出口不可信 / the outlets are not trustworthy
        bError      := TRUE;               // 故障标志置位 / raise the fault flag
        nErrCode    := _nCodeLatch;        // 回放锁存码 / replay the latched code
END_CASE

// 段 8｜步推进后的计时器复位请求（下一拍生效）/ segment 8, request a timer restart after an advance
IF _bAdvanced THEN                         // 本拍发生过推进 / the step advanced this scan
    _bTimerRestart := TRUE;                // 下一拍断 IN 一拍，新步从 0 计时 / drop IN next scan so the new step times from zero
END_IF

// 段 9｜出口映射（名实双出口同源，R191；单点写入，无自赋值）/ segment 9, the outlet mapping
eState  := _eState;                        // 状态出口 = 寄存器 / the state outlet mirrors the register
nStepNo := _nStep;                         // 步号出口 = 寄存器 / the step outlet mirrors the register
END_FUNCTION_BLOCK

(* ---- FB_DL_ReqAckHandshake.st ---- *)
(*
  ==================================================================
  组件名 Component  : FB_DL_ReqAckHandshake
  分类   Category   : DL_Base
  复杂度 Complexity  : 中
  版本   Version    : 1.0.0
  功能   Purpose    : 通用请求-应答握手原子（无工艺语义）。请求上升沿武装进入应答
                      等待相，应答窗 tAck 内收到 bAck 电平则输出确认单拍 bDone；
                      窗到期未见应答则输出重试单拍 bRetry 并进重试间隔相 tRetry，
                      重试次数达 nMaxRetry 仍不应答则锁存故障码。
  来源   Source     : self-std（IEC 61131-3 标准时序语义自研原子）
  溯源   Origin     : 请求-应答握手为公开时序语义，道莅 clean-room 自研实现，
                      未复制任何厂商私有库源码。
  平台   Platform   : 纯 IEC 61131-3（Standard.library: TON / R_TRIG），
                      CODESYS / TwinCAT / InoProShop / Machine Expert 通用
  分工声明 Split     : 与 FB_DL_AgvDockingHandshake（工艺级对接握手）分工——
                      后者承载工位/库位工艺时序与就位判据；本件为无工艺语义的
                      时序原子，只做沿武装、窗超时、重试与锁存，不判任何机械条件。
  作者   Author     : 道莅代码库 · PLC 编程专家（R60）
  ------------------------------------------------------------------
  边界 Boundary     :
                      一 同拍双窗配比约束（R100/R239）：tAck 为单次应答窗、
                         tRetry 为重试间隔，约束 tAck > tRetry > 0——若
                         tRetry >= tAck，重试节拍慢于超时检测，重试上限在等效
                         时间内不可达，重试语义退化为一次性；违反即在段 2
                         组态闸锁存故障码（禁只在注释里声明）；
                      二 单拍输出 bDone / bRetry 统一出口段每拍先预置 FALSE，
                         分支只写 TRUE（R256）；
                      三 首拍零假沿自证（R257）：R_TRIG 内部存储位初值 FALSE，
                         首拍 bReq 已为真即判为一次新请求沿，语义安全（请求电平
                         已存在则握手应立即启动），而 bAck 首拍为真不会误置
                         bDone——它只在应答等待相内被消费；
                      四 应答等待相退出条件三条（R98）：bAck 成立 / 请求撤销
                         （进相前置消失，无码回空闲）/ 应答窗超时；缺一即死等；
                      五 使能 bEnable = FALSE 时语义为「冻结保持 + 弃用请求」
                         （退出活动相回空闲，不锁存、不出单拍）——R191 声明行；
                      六 故障解除路径：eFault 相由复位沿迁回空闲并清锁存与重试
                         计数（bReset 为输入引脚，恒可达，R152 自证）；
                      七 故障码一律锁存回放，不在故障相按当下输入重新推断。
  错误码   Codes    :
    16#0001_0613【故障级】组态非法（窗配比违反或重试上限为负），锁存至复位沿
    16#0001_0614【故障级】应答窗超时且重试耗尽，锁存至复位沿
    16#0001_0615【信息级】重试计数已达上限（本拍为最后一次重试，逐拍重算）
  验收   Acceptance :
    算法已证（脚本）：未跑 ｜ 编译器已证（三平台）：未跑
    V1 tAck=2s、nMaxRetry=2、第 3 个窗到期前给 bAck → bDone 单拍、计数归零
    V2 全程无 bAck、nMaxRetry=2 → 两次 bRetry 单拍后锁码 0614、相冻结
    V3 tRetry >= tAck → 首拍即锁码 0613，无单拍输出
  修订记录 Revision  :
    2026-11-21  v1.0.0  R60 首版（批 1 · 序号 4）
  ==================================================================
*)

TYPE E_DL_ReqAckPhase :
(
    eIdle     := 0,  // 空闲：等请求上升沿或复位 / idle, waiting for the request edge or a reset
    eWaitAck  := 10, // 应答等待：等 bAck / 请求撤销 / 窗超时 / waiting for the acknowledgement, an abort or the window expiry
    eRetryGap := 20, // 重试间隔：等 tRetry 到期后重开应答窗 / the retry gap, reopen the window after tRetry
    eFault    := 30  // 故障：锁存故障码，等复位沿 / fault, the code latched, waiting for the reset edge
);
END_TYPE

FUNCTION_BLOCK FB_DL_ReqAckHandshake
VAR_INPUT
    bEnable    : BOOL := TRUE;  // 使能，FALSE 时退相回空闲（边界五）/ the enable, false returns the phase to idle
    bReq       : BOOL := FALSE; // 请求电平，上升沿武装握手 / the request level, the rising edge arms the handshake
    bAck       : BOOL := FALSE; // 应答电平，仅在应答等待相内被消费 / the acknowledgement level, consumed only inside the waiting phase
    bReset     : BOOL := FALSE; // 复位沿：清故障锁存与重试计数并回空闲 / the reset edge, clears the latch and the retry count then returns to idle
    tAck       : TIME := T#2S;  // 单次应答窗时长 [毫秒] / the single attempt acknowledgement window
    tRetry     : TIME := T#500MS; // 重试间隔时长 [毫秒]，约束 tAck > tRetry / the retry gap, constrained below the window
    nMaxRetry  : DINT := 3;     // 最大重试次数 [次]，域 0..100 / the maximum retry count, from zero to one hundred
END_VAR
VAR_OUTPUT
    bBusy      : BOOL := FALSE;                 // 握手中（等待或重试间隔）[-] / the handshake in progress flag
    bDone      : BOOL := FALSE;                 // 握手成功单拍脉冲 [-] / the success one shot pulse
    bRetry     : BOOL := FALSE;                 // 发起重试单拍脉冲 [-] / the retry one shot pulse
    nRetryCnt  : DINT := 0;                     // 已发起重试次数 [次]，饱和于上限 / the issued retry count, saturated at the bound
    eState     : E_DL_ReqAckPhase;              // 主状态机当前态 [状态] / the current state of the main machine
    bError     : BOOL := FALSE;                 // 故障锁存位 [-] / the latched fault bit
    eErr       : UDINT := 16#0000_0000;         // 错误码，0 = 正常 / the error code, zero is ok
END_VAR
VAR
    _bInit     : BOOL := FALSE;                            // 首拍初始化标志（R310）/ the first scan flag
    _eState    : E_DL_ReqAckPhase := E_DL_ReqAckPhase.eIdle; // 内部状态寄存器，段 3 唯一写点 / the internal state register, single writer
    _nRetryCnt : DINT := 0;                                // 重试计数副本，段 5 单点映射 / the retry count copy, mapped once in segment five
    _bDone     : BOOL := FALSE;                            // 成功单拍内部位，段 1 预清段 5 映射 / the internal success bit, preset then mapped
    _bRetry    : BOOL := FALSE;                            // 重试单拍内部位，段 1 预清段 5 映射 / the internal retry bit, preset then mapped
    _bFault    : BOOL := FALSE;                            // 故障锁存副本（仅复位沿清除）/ the fault latch copy, cleared only on the reset edge
    _bRetrySat : BOOL := FALSE;                            // 重试计数饱和指示（逐拍重算）[-] / the retry saturation flag, recomputed every scan
    _bCfgBad   : BOOL := FALSE;                            // 组态非法指示（逐拍重算）[-] / the configuration fault flag, recomputed every scan
    rtReq      : R_TRIG;                                   // 请求沿实例，段 0 无条件刷新 / the request edge instance, refreshed unconditionally
    rtReset    : R_TRIG;                                   // 复位沿实例，段 0 无条件刷新 / the reset edge instance, refreshed unconditionally
    tonAck     : TON;                                      // 应答窗定时器，段 0 无条件刷新 / the acknowledgement window timer, refreshed unconditionally
    tonRetry   : TON;                                      // 重试间隔定时器，段 0 无条件刷新 / the retry gap timer, refreshed unconditionally
END_VAR
VAR CONSTANT
    DL_RAH_RETRYMAX : DINT := 100; // 重试次数上界 [次]，防组态越域 / the retry count bound against configuration overflow
END_VAR

// 段 0｜定时器与沿检测无条件周期刷新（禁入分支，R7；IN 串故障锁存量门控，FB50-1）/ segment 0, the unconditional refresh with the latch gate
rtReq(CLK := bReq); // 请求沿 / the request edge
rtReset(CLK := bReset); // 复位沿 / the reset edge
tonAck(IN := (_eState = E_DL_ReqAckPhase.eWaitAck) AND (NOT _bFault), PT := tAck); // 应答窗：仅在等待相且无锁存时计时 / the window timing only in the waiting phase without a latch
tonRetry(IN := (_eState = E_DL_ReqAckPhase.eRetryGap) AND (NOT _bFault), PT := tRetry); // 重试间隔计时 / the retry gap timing

// 段 1｜首拍初始化与单拍标志预清（仅单拍标志入清单，R32 FB32-1；R256）/ segment 1, the first scan init and the one shot preset
IF NOT _bInit THEN // 首拍一拍 / the first scan
    _bInit := TRUE; // 置首拍标志 / raise the first scan flag
    _nRetryCnt := 0; // 重试计数显式清零 / clear the retry count explicitly
    _bFault := FALSE; // 故障锁存显式清零 / clear the fault latch explicitly
    _eState := E_DL_ReqAckPhase.eIdle; // 状态显式落空闲 / place the state to idle explicitly
END_IF
_bDone := FALSE; // 成功单拍预清零 / preset the success pulse false
_bRetry := FALSE; // 重试单拍预清零 / preset the retry pulse false
_bRetrySat := FALSE; // 饱和指示预清零 / preset the saturation flag false
_bCfgBad := FALSE; // 组态非法指示预清零 / preset the configuration fault flag false

// 段 2｜组态域闸（窗配比 + 重试上限，边界一；同拍双窗配比在此落成可观测故障）/ segment 2, the configuration gate with the window ratio landed as an observable fault
IF (tAck <= T#0S) OR (tRetry <= T#0S) OR (tRetry >= tAck) OR (nMaxRetry < 0) OR (nMaxRetry > DL_RAH_RETRYMAX) THEN // 任一越域 / any item out of domain
    _bCfgBad := TRUE; // 置组态非法 / raise the configuration fault
    _bFault := TRUE; // 锁存故障（段 4 迁移相）/ latch the fault, the segment four migrates the phase
END_IF

// 段 3｜主状态机（ENUM + CASE，ELSE 拦非法态）/ segment 3, the main machine with the illegal state guard
CASE _eState OF
    E_DL_ReqAckPhase.eIdle: // 空闲相：等请求沿 / the idle phase, waiting for the request edge
        IF bEnable AND (NOT _bFault) AND rtReq.Q THEN // 迁入判据：使能且无锁存且有请求沿（R274 全量闸位复检）/ the entry with the full gate recheck
            _nRetryCnt := 0; // 新一轮握手重试计数归零 / reset the retry count for the new round
            _eState := E_DL_ReqAckPhase.eWaitAck; // 迁入应答等待相 / enter the waiting phase
        END_IF
    E_DL_ReqAckPhase.eWaitAck: // 应答等待相：三条退出（边界四，R98）/ the waiting phase with three exits
        IF bAck THEN // 出口一：应答成立 / the first exit, the acknowledgement
            _bDone := TRUE; // 置成功单拍 / raise the success pulse
            _nRetryCnt := 0; // 成功后计数归零（复位作用域：清累计量）/ on success the count returns to zero
            _eState := E_DL_ReqAckPhase.eIdle; // 迁回空闲 / back to idle
        ELSIF (NOT bReq) THEN // 出口二：请求撤销（进相前置条件已消失，无码回空闲）/ the second exit, the request withdrawn with no code
            _nRetryCnt := 0; // 计数归零 / the count returns to zero
            _eState := E_DL_ReqAckPhase.eIdle; // 迁回空闲 / back to idle
        ELSIF tonAck.Q THEN // 出口三：应答窗到期 / the third exit, the window expired
            IF _nRetryCnt < nMaxRetry THEN // 尚有重试额度 / a retry remains available
                _nRetryCnt := _nRetryCnt + 1; // 重试计数推进 / advance the retry count
                _bRetry := TRUE; // 置重试单拍 / raise the retry pulse
                IF _nRetryCnt >= nMaxRetry THEN // 已用尽全部额度 / the whole allowance is used
                    _bRetrySat := TRUE; // 置饱和提示（最后一次重试，信息级）/ raise the informational saturation hint
                END_IF
                _eState := E_DL_ReqAckPhase.eRetryGap; // 迁入重试间隔相 / enter the retry gap phase
            ELSE // 额度已尽 / the allowance exhausted
                _bFault := TRUE; // 锁存故障（0614，段 4 迁移相）/ latch the fault, migrated in segment four
            END_IF
        END_IF
        IF (_eState = E_DL_ReqAckPhase.eWaitAck) AND (NOT bEnable) AND (NOT _bFault) THEN // 失能弃用请求（不借故障相过桥，R211；相判据防成功拍被改写）/ the disable discards the request without bridging the fault phase
            _nRetryCnt := 0; // 计数归零 / the count returns to zero
            _eState := E_DL_ReqAckPhase.eIdle; // 迁回空闲 / back to idle
        END_IF
    E_DL_ReqAckPhase.eRetryGap: // 重试间隔相：等间隔到期或请求撤销 / the retry gap phase
        IF (NOT bReq) THEN // 退出条件一：请求撤销（前置消失）/ the first exit, the request withdrawn
            _nRetryCnt := 0; // 计数归零 / the count returns to zero
            _eState := E_DL_ReqAckPhase.eIdle; // 迁回空闲 / back to idle
        ELSIF tonRetry.Q THEN // 退出条件二：间隔到期，重开应答窗 / the second exit, the gap expired, reopen the window
            _eState := E_DL_ReqAckPhase.eWaitAck; // 迁回应答等待相 / back to the waiting phase
        END_IF
        IF (NOT bEnable) AND (NOT _bFault) THEN // 失能回空闲 / the disable returns to idle
            _nRetryCnt := 0; // 计数归零 / the count returns to zero
            _eState := E_DL_ReqAckPhase.eIdle; // 迁回空闲 / back to idle
        END_IF
    E_DL_ReqAckPhase.eFault: // 故障相：锁存保持，等复位沿（解除路径可达，边界六）/ the fault phase, held until the reset edge
        IF rtReset.Q THEN // 复位沿（复位作用域：清锁存 + 清累计量 + 迁相位）/ the reset edge with the declared scope
            _bFault := FALSE; // 清故障锁存 / clear the fault latch
            _nRetryCnt := 0; // 清重试计数 / clear the retry count
            _eState := E_DL_ReqAckPhase.eIdle; // 故障相迁出边回空闲 / the exit edge back to idle
        END_IF
    ELSE // 非法枚举值拦截 / the illegal enumeration guard
        _eState := E_DL_ReqAckPhase.eIdle; // 落回空闲 / force back to idle
        _bFault := TRUE; // 置故障锁存 / latch the fault
END_CASE

// 段 4｜故障锁存迁移闸（置于解除段之后防同拍抢迁，R258）/ segment 4, the fault latch to phase gate placed after the release
IF _bFault AND (_eState <> E_DL_ReqAckPhase.eFault) THEN // 已锁存但不在故障相 / latched but not in the fault phase
    _eState := E_DL_ReqAckPhase.eFault; // 迁入故障相 / enter the fault phase
END_IF

// 段 5｜统一出口（内部副本单点映射，R180；故障码锁存回放，R187）/ segment 5, the unified outlet
bBusy := (_eState = E_DL_ReqAckPhase.eWaitAck) OR (_eState = E_DL_ReqAckPhase.eRetryGap); // 握手中指示 / the in progress flag
bDone := _bDone; // 成功单拍出口 / the success pulse outlet
bRetry := _bRetry; // 重试单拍出口 / the retry pulse outlet
nRetryCnt := _nRetryCnt; // 重试计数出口 / the retry count outlet
eState := _eState; // 状态出口 / the state outlet
bError := _bFault; // 故障位出口（与锁存同源）/ the fault bit outlet from the same latch
IF _bFault THEN // 故障锁存回放优先 / the latched fault replays first
    IF _bCfgBad THEN // 组态成因 / the configuration cause
        eErr := 16#0001_0613; // 故障级：组态非法 / fault grade, the configuration is illegal
    ELSE // 超时成因（独立码值，R190 归因唯一）/ the timeout cause with its own code value
        eErr := 16#0001_0614; // 故障级：应答窗超时且重试耗尽 / fault grade, the window expired with the retries exhausted
    END_IF
ELSIF _bRetrySat THEN // 信息级提示 / the informational hint
    eErr := 16#0001_0615; // 信息级：重试计数已达上限 / informational, the retry count reached the bound
ELSE // 无事件 / no event
    eErr := 16#0000_0000; // 正常 / ok
END_IF
END_FUNCTION_BLOCK

(* ---- FB_DL_RolloverCounterUdint.st ---- *)
(*
  ==================================================================
  组件名 Component  : FB_DL_RolloverCounterUdint
  分类   Category   : DL_Base
  复杂度 Complexity  : 中
  版本   Version    : 1.0.0
  功能   Purpose    : UDINT 域回绕计数器。计数沿推进，计数达回绕上限 uUpper 后
                      下一沿回到 0 并出回绕单拍脉冲 bRoll，圈数 nTurns 累计并饱和；
                      装载电平优先于计数沿；上限非法（0）时退化冻结并锁存故障码。
  来源   Source     : t2-1-lgf-counter（LGF Counter 回绕计数族 UDINT 变体）
  溯源   Origin     : 回绕计数属公开计数语义，clean-room 自研实现，未复制 LGF
                      或任何厂商私有库源码。
  平台   Platform   : 纯 IEC 61131-3（TON 未用；仅 R_TRIG / FOR 无关；无位运算），
                      CODESYS / TwinCAT / InoProShop / Machine Expert 通用
  分工声明 Split     : 与 FB_DL_RolloverCounter（INT 属主）与 FB_DL_ModuloCounter
                      （取模索引属主）三角互引——本件为 UDINT 域回绕计数，
                      只出计数/圈数/回绕脉冲，不做取模索引换算、不做工艺计件。
                      INT 属主仍管有符号双向回绕，本件不接管负向语义。
  作者   Author     : 道莅代码库 · PLC 编程专家（R60）
  ------------------------------------------------------------------
  边界 Boundary     :
                      一 回绕一律「比较 + 赋值」，禁用 MOD（负数取余三平台歧义）：
                         自增前判 uCount >= uUpper，命中则置 0 并计一圈；
                      二 整数进位点自证：uUpper=59 时计数序列 …58→59→0 圈数 +1；
                         uUpper=0 判非法冻结（不成环，禁静默计成 0 长循环）；
                      三 自增域自证：仅在 uCount < uUpper 时执行 +1，而
                         uUpper <= 16#FFFF_FFFF，故不存在 16#FFFF_FFFF + 1 回绕；
                      四 装载 bLoad 电平优先于复位沿与计数沿；装载值超上限钳位；
                      五 使能 bEnable = FALSE 时语义为「冻结保持」（计数/圈数/
                         回绕脉冲均保持，本拍不出脉冲）——本条为 R191 声明行；
                      六 故障解除路径：上限恢复合法（uUpper >= 1）且复位沿到达，
                         故障相迁回 eIdle 并清锁存（R152 可达性自证：uUpper 为
                         输入引脚，可恒达）。
  接口偏离声明       : 派单示意 nPreset（有符号命名），UDINT 域按 R265 命名-类型
                      一致性落为 uPreset，语义一字不减。
  错误码   Codes    :
    16#0001_0610【信息级】装载值或现存计数超上限已钳位（同一语义共码，R90 反证：
                         二者都只由「钳到 uUpper」观测，无独立可观测差异，不加第 4 码）
    16#0001_0611【信息级】圈数已饱和（达 DINT 计数上限，停止累计）
    16#0001_0612【故障级】回绕上限非法（0），计数退化冻结（锁存至复位沿）
  验收   Acceptance :
    算法已证（脚本）：未跑 ｜ 编译器已证（三平台）：未跑
    V1 uUpper=59，连打 60 沿 → 第 60 沿后 uCount=0、nTurns=1、bRoll 单拍
    V2 uUpper=0 → eFrozen、码 0612、bError 锁存，计数保持
    V3 bLoad 与 bCount 同拍 → 装载优先，计数等于钳位后的 uPreset
  修订记录 Revision  :
    2026-11-21  v1.0.0  R60 首版（批 1 · 序号 3）
  ==================================================================
*)

TYPE E_DL_RolloverPhaseUd :
(
    eIdle   := 0,  // 空闲：未使能，计数与圈数保持 / idle, disabled, the count and the turns held
    eCount  := 10, // 计数：按装载与计数沿推进并回绕 / counting, driven by the load and the count edges with wrap around
    eFrozen := 20  // 冻结：上限非法，计数保持并报警 / frozen, the bound is illegal, the count held with the alarm
);
END_TYPE

FUNCTION_BLOCK FB_DL_RolloverCounterUdint
VAR_INPUT
    bEnable    : BOOL;  // 使能，FALSE 时冻结保持（边界五）/ the enable, false freezes and holds
    bReset     : BOOL;  // 复位上升沿：计数与圈数清零 / the reset rising edge, clears the count and the turns
    bCount     : BOOL;  // 计数上升沿：计数推进或回绕 / the count rising edge, advance or wrap
    bLoad      : BOOL;  // 装载电平，优先级最高（边界四）/ the level true load, the highest priority
    uPreset    : UDINT; // 装载预置值 [计数值]，超上限时钳位 / the load preset, clamped to the bound
    uUpper     : UDINT; // 回绕上限（含）[计数值]，合法域 1..16#FFFF_FFFF / the wrap bound inclusive, legal from one to the unsigned maximum
END_VAR
VAR_OUTPUT
    uCount    : UDINT;                  // 当前计数值 [计数值]，域 0..uUpper / the current count, from zero to the bound
    bRoll     : BOOL;                   // 本拍回绕单拍脉冲 [-] / the wrap one shot pulse of this scan
    nTurns    : DINT;                   // 累计圈数（饱和）[圈] / the accumulated turns, saturated
    bAtUpper  : BOOL;                   // 当前值已达回绕上限（逐拍重算）[-] / the count reached the bound, recomputed every scan
    eState    : E_DL_RolloverPhaseUd;   // 主状态机当前态 [状态] / the current state of the main machine
    bError    : BOOL;                   // 故障锁存位 [-] / the latched fault bit
    eErr      : UDINT;                  // 错误码，0 = 正常 / the error code, zero is ok
END_VAR
VAR
    _bInit     : BOOL := FALSE;                  // 首拍初始化标志（R310）/ the first scan flag
    _eState    : E_DL_RolloverPhaseUd := E_DL_RolloverPhaseUd.eIdle; // 内部状态寄存器，段 3 唯一写点 / the internal state register, single writer
    _uCount    : UDINT := 0;                     // 计数内部副本，段 5 单点映射 / the internal count copy, mapped once in segment five
    _nTurns    : DINT := 0;                      // 圈数内部副本，段 5 单点映射 / the internal turns copy, mapped once in segment five
    _bRoll     : BOOL := FALSE;                  // 回绕单拍内部位，段 1 预清段 5 映射 / the internal wrap pulse bit, preset then mapped
    _bFault    : BOOL := FALSE;                  // 故障锁存副本（仅复位沿清除）/ the fault latch copy, cleared only on the reset edge
    _bTurnSat  : BOOL := FALSE;                  // 圈数饱和指示（逐拍重算）[-] / the turn saturation flag, recomputed every scan
    _bClamped  : BOOL := FALSE;                  // 钳位事件标记（逐拍重算）[-] / the clamp event flag, recomputed every scan
    rtCount    : R_TRIG;                         // 计数沿实例，段 0 无条件刷新 / the count edge instance, refreshed unconditionally
    rtReset    : R_TRIG;                         // 复位沿实例，段 0 无条件刷新 / the reset edge instance, refreshed unconditionally
END_VAR
VAR CONSTANT
    DL_RCU_TURNMAX : DINT := 1000000000; // 圈数饱和上界 [圈]，留足 INT 域余量防溢出 / the turn saturation bound with margin against overflow
END_VAR

// 段 0｜沿检测无条件周期刷新（禁入分支，R7）；本件无 TON / segment 0, the unconditional edge refresh
rtCount(CLK := bCount); // 计数沿 / the count edge
rtReset(CLK := bReset); // 复位沿 / the reset edge

// 段 1｜首拍初始化与单拍标志预清（单拍标志入清单，保持型量不入，R32 FB32-1）/ segment 1, the first scan init and the one shot preset
IF NOT _bInit THEN // 首拍一拍 / the first scan
    _bInit := TRUE; // 置首拍标志 / raise the first scan flag
    _uCount := 0; // 计数显式清零 / clear the count explicitly
    _nTurns := 0; // 圈数显式清零 / clear the turns explicitly
    _bFault := FALSE; // 故障锁存显式清零 / clear the fault latch explicitly
    _eState := E_DL_RolloverPhaseUd.eIdle; // 状态显式落空闲 / place the state to idle explicitly
END_IF
_bRoll := FALSE; // 回绕脉冲预清零（先清后置，段 3 只写 TRUE）/ preset the wrap pulse false, the segment three only raises it
_bTurnSat := FALSE; // 饱和指示预清零 / preset the saturation flag false
_bClamped := FALSE; // 钳位标记预清零 / preset the clamp flag false

// 段 2｜组态域闸与钳位（上限非法 → 故障锁存；装载值/现存计数超上限 → 钳位，边界二四）/ segment 2, the configuration gate and the clamps
IF uUpper < 1 THEN // 上限非法：不成环 / an illegal bound, no ring exists
    _bFault := TRUE; // 锁存故障（段 4 迁移相）/ latch the fault, the segment four migrates the phase
ELSE // 上限合法：施加钳位 / a legal bound, apply the clamps
    IF uPreset > uUpper THEN // 装载值超上限 / the load preset above the bound
        _bClamped := TRUE; // 记钳位事件 / register the clamp event
    END_IF
    IF _uCount > uUpper THEN // 上限在线改小致现存计数越界（边界二回钳）/ the bound reduced online puts the count above it
        _uCount := uUpper; // 现存计数回钳（回钳后不再复判越界，R241）/ clamp the count back, no re-test afterwards
        _bClamped := TRUE; // 记钳位事件 / register the clamp event
    END_IF
END_IF

// 段 3｜主状态机（ENUM + CASE，ELSE 拦非法态）/ segment 3, the main machine with the illegal state guard
CASE _eState OF
    E_DL_RolloverPhaseUd.eIdle: // 空闲相：未使能或已复位 / the idle phase, disabled or reset
        IF bReset AND rtReset.Q THEN // 复位沿（空闲相也清零，复位作用域：清累计量）/ the reset edge, the scope is the accumulated quantity
            _uCount := 0; // 计数清零 / clear the count
            _nTurns := 0; // 圈数清零 / clear the turns
        END_IF
        IF bEnable AND (_bFault = FALSE) AND (uUpper >= 1) THEN // 迁入条件：使能且无故障且上限合法（R274 全量闸位复检）/ the entry with the full gate recheck
            _eState := E_DL_RolloverPhaseUd.eCount; // 迁入计数相 / enter the counting phase
        END_IF
    E_DL_RolloverPhaseUd.eCount: // 计数相：装载优先，其次计数沿，再次复位沿 / the counting phase, load first, then the count edge, then the reset edge
        IF bLoad THEN // 装载电平优先（边界四）/ the load level wins
            IF uPreset > uUpper THEN // 装载值超上限 / the preset above the bound
                _uCount := uUpper; // 钳到上限 / clamp to the bound
            ELSE // 装载值域内 / the preset inside the domain
                _uCount := uPreset; // 直接装载 / take the preset
            END_IF
        ELSIF rtCount.Q THEN // 计数沿：自增前判回绕（边界一三）/ the count edge, test the wrap before the increment
            IF _uCount >= uUpper THEN // 已达上限，本沿回绕 / at the bound, wrap on this edge
                _uCount := 0; // 回绕置零 / wrap to zero
                _bRoll := TRUE; // 置回绕单拍 / raise the wrap pulse
                IF _nTurns < DL_RCU_TURNMAX THEN // 圈数未饱和 / the turns not saturated
                    _nTurns := _nTurns + 1; // 圈数推进 / advance the turns
                ELSE // 圈数饱和 / the turns saturated
                    _bTurnSat := TRUE; // 置饱和指示 / raise the saturation flag
                END_IF
            ELSE // 未达上限，正常自增（不存在位型回绕）/ below the bound, a plain increment with no bit pattern wrap
                _uCount := _uCount + 1; // 计数自增 / advance the count
            END_IF
        ELSIF bReset AND rtReset.Q THEN // 复位沿（复位作用域：清累计量 + 清回绕脉冲由段 1 预清承担）/ the reset edge
            _uCount := 0; // 计数清零 / clear the count
            _nTurns := 0; // 圈数清零 / clear the turns
        END_IF
        IF (NOT bEnable) AND (_bFault = FALSE) THEN // 失能回空闲（不借故障相过桥，R211）/ disable returns to idle without bridging the fault phase
            _eState := E_DL_RolloverPhaseUd.eIdle; // 迁回空闲 / back to idle
        END_IF
    E_DL_RolloverPhaseUd.eFrozen: // 冻结相：上限非法，计数保持 / the frozen phase, illegal bound, the count held
        IF rtReset.Q AND (uUpper >= 1) THEN // 解除式：复位沿且上限已恢复合法（R152 可达）/ the release, a reset edge with a legal bound restored
            _bFault := FALSE; // 清故障锁存 / clear the fault latch
            _uCount := 0; // 复位作用域：清累计量 / the reset scope, clear the accumulated quantity
            _nTurns := 0; // 复位作用域：清累计量 / the reset scope, clear the accumulated quantity
            _eState := E_DL_RolloverPhaseUd.eIdle; // 故障相迁出边（迁回空闲）/ the exit edge back to idle
        END_IF
    ELSE // 非法枚举值拦截 / the illegal enumeration guard
        _eState := E_DL_RolloverPhaseUd.eIdle; // 落回空闲 / force back to idle
        _bFault := TRUE; // 置故障锁存 / latch the fault
END_CASE

// 段 4｜故障锁存迁移闸（置于解除段之后，R258；锁存即迁冻结相）/ segment 4, the fault latch to phase gate, placed after the release
IF _bFault AND (_eState <> E_DL_RolloverPhaseUd.eFrozen) THEN // 已锁存但未在冻结相 / latched but not in the frozen phase
    _eState := E_DL_RolloverPhaseUd.eFrozen; // 迁入冻结相 / enter the frozen phase
END_IF

// 段 5｜统一出口（内部副本单点映射，R180；故障码锁存回放，R187）/ segment 5, the unified outlet
uCount := _uCount; // 计数出口 / the count outlet
nTurns := _nTurns; // 圈数出口 / the turns outlet
bRoll := _bRoll; // 回绕单拍出口 / the wrap pulse outlet
bAtUpper := (_uCount >= uUpper) AND (uUpper >= 1); // 达上限指示（上限非法时不宣称，逐拍重算）/ the at bound flag, recomputed every scan
eState := _eState; // 状态出口 / the state outlet
bError := _bFault; // 故障位出口（与锁存同源）/ the fault bit outlet from the same latch
IF _bFault THEN // 故障锁存回放优先 / the latched fault replays first
    eErr := 16#0001_0612; // 故障级：回绕上限非法，计数退化冻结 / fault grade, the illegal bound with the frozen count
ELSIF _bClamped THEN // 其次钳位信息级 / then the clamp informational code
    eErr := 16#0001_0610; // 信息级：超上限已钳位 / informational, clamped to the bound
ELSIF _bTurnSat THEN // 再次圈数饱和信息级 / then the saturation informational code
    eErr := 16#0001_0611; // 信息级：圈数已饱和 / informational, the turns saturated
ELSE // 无事件 / no event
    eErr := 16#0000_0000; // 正常 / ok
END_IF
END_FUNCTION_BLOCK

(* ---- FB_DL_RSBistable.st ---- *)
(*==============================================================================
 * 组件名称 (Component)  : FB_DL_RSBistable
 * 所属子库 (Sublibrary) : DL_Base
 * 当前版本 (Version)    : 1.0.0
 * 兼容性   (Platform)   : CODESYS 3.5 / TwinCAT 3 / 汇川 InoProShop / Machine Expert
 *                         仅依赖纯 IEC 61131-3 标准运算符，零厂商方言
 * 功能描述 (Function)   : RS 复位优先双稳态防御包装。内部委托 IEC 61131-3 标准
 *                         RS 语义（bQ := (bS OR bQ) AND NOT bR1），外围提供
 *                         S/R1 同拍仲裁显式化与仲裁诊断码输出。
 *                         与 FB_DL_SRBistable 为镜像件（SR=置位优先，RS=复位优先），
 *                         选型时以"同拍竞态时谁说了算"为准，两者头注释互引。
 * 溯源     (Origin)     : IEC 61131-3 标准语义的道莅防御性实现
 *                         （接口语义由 IEC 61131-3 定义，clean-room 重写，
 *                         参考公开标准条款）
 * 码位     (Diag Codes) : 信息级占用区间 16#0001_014E（本件独占，仅此一码）
 *                         16#0001_014E = S/R1 同拍为 TRUE，复位胜出（标准语义，
 *                         仅供现场排查，不置故障）
 * 类型裁定 (Type Note)  : 码位段 16#0001_xxxx 为全库共享 32 位段，WORD 容量不足，
 *                         故 uDiag 采用 UDINT 承载（与库内 uErrorId : UDINT 惯例一致）
 * 依赖     (Depends)    : 无 DL_ 内部依赖；无标准库实例（纯布尔逻辑）
 * 红线自检 (Redline)    : R1 ✓ 零全局变量与外部变量引用 ｜ R2 ✓ 零物理 IO 地址直写
 *                         R3 ✓ 纯 IEC 61131-3 ｜ R4 ✓ 同拍仲裁显式化+首扫初始化
 *                         R5 ✓ 全变量中英双语同行注释 ｜ R6 N/A（无顺序状态机，见下）
 *                         R7 ✓ 无定时器/沿检测实例（N/A）
 * 说明     (Note)       : R6 标注 N/A —— 本组件为组合逻辑双稳态，不存在顺序状态机，
 *                         无 CASE 可写；非法状态不可能出现（唯一状态即输出锁存），
 *                         故以本节说明替代 ELSE 兜底，符合"无状态机则标注 N/A"口径。
 * 防御行为声明 (Defense): ① S 与 R1 同拍为 TRUE 时按 IEC 语义复位优先（R1 胜出），
 *                           同时置信息级诊断码 16#0001_014E，下拍仲裁消失自动清零；
 *                         ② 首扫输出初始化为 FALSE，杜绝上电假输出。
 * 修订历史 (Revision)   :
 *   2026-11-16  v1.0.0  首版入库（R14 批 1 · T0 快车道）
 *============================================================================*)
FUNCTION_BLOCK FB_DL_RSBistable
VAR_INPUT
    bS  : BOOL;  // 置位输入，仅在 R1 为 FALSE 的拍次生效 / Set input, effective only on scans where R1 is FALSE
    bR1 : BOOL;  // 复位主导输入（IEC R1 语义），TRUE 时输出无条件复位 / Reset-dominant input (IEC R1), TRUE forces output reset
END_VAR
VAR_OUTPUT
    bQ    : BOOL;   // 复位优先输出（IEC Q1 语义），TRUE 保持至复位 / Reset-dominant output (IEC Q1), latched TRUE until reset
    uDiag : UDINT;  // 仲裁诊断字，16#0001_014E=S/R1 同拍复位胜出，0=无仲裁事件 / Arbitration diag word, 16#0001_014E=same-scan S/R1 with reset winning, 0=no arbitration
END_VAR
VAR
    xInit : BOOL;   // 首扫初始化标志，FALSE=尚未完成上电初始化 / First-scan init flag, FALSE = power-on init not yet done
END_VAR

(*------------------------------------------------------------------------------
 * 段 1｜首扫初始化（历史教训⑤口径）：置于逻辑最前，禁止"初值置位后同步清零"反模式
 *      First-scan init (lesson 5): placed at the very front of the logic body
 *-----------------------------------------------------------------------------*)
IF NOT xInit THEN
    xInit := TRUE;      // 置初始化完成标志 / Mark init as done
    bQ    := FALSE;     // 首扫输出强制 FALSE，杜绝上电假输出 / Force output FALSE on first scan
    uDiag := 16#0000_0000;  // 首扫诊断字清零 / Clear diag word on first scan
END_IF

(*------------------------------------------------------------------------------
 * 段 2｜同拍仲裁诊断：S 与 R1 同拍为 TRUE 是标准定义的合法竞态，置信息码不置故障
 *      Same-scan arbitration diag: S AND R1 is a legal race per the standard,
 *      informational code only, never a fault
 *-----------------------------------------------------------------------------*)
IF bS AND bR1 THEN
    uDiag := 16#0001_014E;  // 同拍竞态：复位优先胜出（信息级）/ Same-scan race: reset-dominant wins (informational)
ELSE
    uDiag := 16#0000_0000;  // 无竞态，诊断字清零 / No race, clear diag word
END_IF

(*------------------------------------------------------------------------------
 * 段 3｜RS 复位优先核心语义（委托 IEC 61131-3 标准 RS 定义，不重实现）：
 *      bQ := (bS OR bQ) AND NOT bR1，右侧 bQ 取上一拍锁存值
 *      RS reset-dominant core semantics (delegates to the IEC 61131-3 RS definition);
 *      the bQ on the right-hand side reads the latched value of the previous scan
 *-----------------------------------------------------------------------------*)
bQ := (bS OR bQ) AND NOT bR1;  // 复位优先：R1=1 恒复位，R1=0 且 S=1 才置位 / Reset-dominant: R1=1 always resets, set only when R1=0 and S=1
END_FUNCTION_BLOCK

(* ---- FB_DL_RsEx.st ---- *)
(*==============================================================================
 * 组件名称 (Component)  : FB_DL_RsEx
 * 所属子库 (Sublibrary) : DL_Base
 * 当前版本 (Version)    : 1.0.0
 * 兼容性   (Platform)   : CODESYS 3.5 / TwinCAT 3 / 汇川 InoProShop / Machine Expert
 *                         仅依赖纯 IEC 61131-3 标准运算符，零厂商方言
 * 功能描述 (Function)   : RS 复位优先双稳态防御包装。内部委托 IEC 61131-3 标准
 *                         RS 语义（bQ1 := (NOT bR1) AND (bS OR bQ1)），外围提供
 *                         S/R1 同拍仲裁显式化诊断与主从双输出镜像。
 * 溯源     (Origin)     : IEC 61131-3 标准语义的道莅防御性实现
 *                         （接口语义由 IEC 61131-3 定义，clean-room 重写，
 *                         参考公开标准条款，未复制任何闭源厂商源码）
 * 码位     (Diag Codes) : 信息级占用区间 16#0001_049B（本件独占，仅此一码）
 *                         16#0001_049B = S/R1 同拍为 TRUE，复位胜出（标准语义，
 *                         仅供现场排查，不置故障）
 *                         （R90 反证句：同拍仲裁事实无法由 bQ1 观测——复位胜出与
 *                           单纯复位的输出同为 FALSE，现有输出组合无法还原「曾发生
 *                           同拍竞争」，故占信息码）
 * 类型裁定 (Type Note)  : 码位段 16#0001_xxxx 为全库共享 32 位段，WORD 容量不足，
 *                         故 uDiag 采用 UDINT 承载（与库内 uErrorId : UDINT 惯例一致）
 * 依赖     (Depends)    : 无 DL_ 内部依赖；无标准库实例（纯布尔逻辑）
 * 对偶声明 (Dual Note)  : 本件与 FB_DL_SrEx 严格对偶（仲裁优先级互逆：SR 置位优先、
 *                         RS 复位优先；注释结构逐条对照，仲裁语义方向相反）。
 * 红线自检 (Redline)    : R1 ✓ 零全局变量与外部变量引用 ｜ R2 ✓ 零物理 IO 地址直写
 *                         R3 ✓ 纯 IEC 61131-3 ｜ R4 ✓ 同拍仲裁显式化，无浮点无除法
 *                         R5 ✓ 全变量中英双语同行注释 ｜ R6 N/A（无顺序状态机，见下）
 *                         R7 N/A 无定时器与沿检测实例（纯组合保持逻辑）
 * 说明     (Note)       : R6 标注 N/A —— 本组件为单步双稳态保持逻辑，不存在顺序
 *                         状态机，无 CASE 可写；非法状态不可能出现（唯一状态即
 *                         「保持 / 置位 / 复位」三态组合，由标准布尔语义全覆盖），
 *                         故以本节说明替代 ELSE 兜底，符合"无状态机则标注 N/A"口径。
 * 输出语义声明 (R191)   : bS = FALSE 且 bR1 = FALSE 时输出保持末值（双稳态记忆语义），
 *                         非降级非冻结，由标准 RS 语义保证；主从输出 bQ1 与 bQ1M
 *                         单点同源赋值（名实双出口，R191 名实相符）。
 * 修订历史 (Revision)   :
 *   2026-11-19  v1.0.0  首版入库（R40 批 4 · T0 快车道）
 *============================================================================*)
FUNCTION_BLOCK FB_DL_RsEx
VAR_INPUT
    bS  : BOOL;  // 置位输入，TRUE 请求置位，与复位同拍时被复位优先压制 ｜ set input, TRUE requests set, suppressed when simultaneous with the reset
    bR1 : BOOL;  // 复位输入，TRUE 请求复位，与置位同拍时复位优先胜出 ｜ reset input, TRUE requests reset, wins the arbitration when simultaneous with the set
END_VAR
VAR_OUTPUT
    bQ1   : BOOL;  // 主输出，复位优先双稳态 ｜ main output of the reset-dominant bistable
    bQ1M  : BOOL;  // 从输出，与 bQ1 同源镜像（名实双出口）｜ mirror output, same source as bQ1
    uDiag : UDINT; // 诊断字，16#0001_049B=S/R1 同拍复位胜出，0=无诊断事件 ｜ diag word, 16#0001_049B=reset wins on simultaneous S/R1, 0=no diag event
END_VAR

// 段 1｜RS 复位优先标准语义主体（IEC 61131-3 双稳态，不重实现状态内核） ｜ RS reset-dominant standard semantics (IEC 61131-3 bistable, no kernel re-implementation)
bQ1 := (NOT bR1) AND (bS OR bQ1); // 复位优先：R1 为真复位，S 单独为真置位，同拍复位胜出 ｜ reset-dominant: R1 resets, S alone sets, the reset wins on simultaneity

// 段 2｜同拍仲裁显式化诊断（信息级每拍重算口径） ｜ simultaneous-arbitration diagnostics (info level, recomputed every scan)
IF bS AND bR1 THEN
    uDiag := 16#0001_049B; // 同拍仲裁：复位优先胜出（信息级，仅排查用）｜ simultaneous arbitration: the reset wins (info level, for troubleshooting only)
ELSE
    uDiag := 16#0000_0000; // 无同拍仲裁事件，清码（信息级允许每拍重算）｜ no arbitration event, clear the code (info level may be recomputed per scan)
END_IF

// 段 3｜主从输出镜像：单点同源赋值（R191 名实双出口） ｜ main-mirror output: single same-source assignment (R191 paired exits)
bQ1M := bQ1; // 从输出镜像主输出 ｜ the mirror output copies the main output
END_FUNCTION_BLOCK

(* ---- FB_DL_RtoEx.st ---- *)
(*==============================================================================
 * 组件名称 (Component)  : FB_DL_RtoEx
 * 所属子库 (Sublibrary) : DL_Base
 * 当前版本 (Version)    : 1.0.0
 * 兼容性   (Platform)   : CODESYS 3.5 / TwinCAT 3 / 汇川 InoProShop / Machine Expert
 *                         仅依赖 Standard.library（TON），零厂商方言
 * 功能描述 (Function)   : 保持型（累加）定时器防御包装。IEC 61131-3 无标准 RTO
 *                         块，本件按通用 RTO 语义以「内建 TON + 内部累加状态位」
 *                         实现：bIN 断开时冻结累计值（掉保持），bIN 恢复后续计，
 *                         bRESET 任意时刻清零累计（复位优先级最高）。
 * 溯源     (Origin)     : IEC 61131-3 标准语义的道莅防御性实现
 *                         （RTO 非标准块，按通用 RTO 语义 clean-room 实现，
 *                         计时内核委托内建 TON，重实现最小化）
 * 码位     (Diag Codes) : 信息级占用区间 16#0001_0152（本件独占，仅此一码）
 *                         16#0001_0152 = tPT 为负值，已钳位为 T#0s（信息级，
 *                         钳位属正常防御行为，不置故障）
 * 类型裁定 (Type Note)  : 码位段 16#0001_xxxx 为全库共享 32 位段，WORD 容量不足，
 *                         故 uDiag 采用 UDINT 承载（与库内 uErrorId : UDINT 惯例一致）
 * 依赖     (Depends)    : 无 DL_ 内部依赖；Standard.library: TON
 * 红线自检 (Redline)    : R1 ✓ 零全局变量与外部变量引用 ｜ R2 ✓ 零物理 IO 地址直写
 *                         R3 ✓ 纯 IEC 61131-3 ｜ R4 ✓ PT 钳位+越界无涉（纯时间加法）
 *                         R5 ✓ 全变量中英双语同行注释 ｜ R6 N/A（无顺序状态机，见下）
 *                         R7 ✓ TON 实例主体无条件周期刷新
 * 说明     (Note)       : R6 标注 N/A —— 本组件为「使能/暂停/复位」三态时序逻辑，
 *                         非顺序步进状态机，无 CASE 可写；三态互斥由优先级链
 *                         （复位 > 使能）显式保证，无非法态可陷入，以本节说明
 *                         替代 ELSE 兜底，符合"无状态机则标注 N/A"口径。
 * 防御行为声明 (Defense): ① tPT < T#0s 时钳位为 T#0s 并置信息码 16#0001_0152；
 *                         ② 优先级链写死：bRESET（电平）> bIN 使能，复位拍即使
 *                           bIN=TRUE 也清零并重新计时（RTO 通用语义）；
 *                         ③ 掉保持/恢复语义：bIN 断开当拍，上一扫描周期的实时
 *                           计时值被冻结累入保持量（tETLast 在内建 TON 被本次
 *                           调用清零前取用），bIN 恢复后从保持量续计，tET 只增
 *                           不减直至复位；
 *                         ④ 计时中途变更 tPT：以完成时刻的 PT 值计入保持量，
 *                           语义为"以完成时刻预置为准"，头注释留档；
 *                         ⑤ tPT 钳 0（含负钳 0）时 bQ 上电使能即到时（ET>=PT
 *                           恒真），属正常防御行为；
 *                         ⑥ 内部状态量写入点排序审计（历史教训⑦）：复位类
 *                           写入（清累计/清到时位）前置，置位类写入（冻结累加/
 *                           到时锁存）后置，复位沿不被吞。
 * 修订历史 (Revision)   :
 *   2026-11-16  v1.0.0  首版入库（R14 批 2 · T0 快车道）
 *============================================================================*)
FUNCTION_BLOCK FB_DL_RtoEx
VAR_INPUT
    bIN    : BOOL;  // 计时使能，TRUE 累计计时，FALSE 暂停并保持累计值 / Timing enable, TRUE accumulates, FALSE pauses and holds the accumulated time
    bRESET : BOOL;  // 复位输入（电平，优先级最高），清零累计与到时位 / Reset input (level, highest priority), clears accumulation and done flag
    tPT    : TIME;  // 预置总延时 [ms]，负值将被钳位为 T#0s / Preset total delay [ms], negative values are clamped to T#0s
END_VAR
VAR_OUTPUT
    bQ    : BOOL;   // 累计到达输出，累计值达 tPT 后保持 / Accumulated-done output, held TRUE once accumulation reaches tPT
    tET   : TIME;   // 累计值 [ms]，bIN 断开保持、只增不减至复位 / Accumulated time [ms], held on bIN drop, only grows until reset
    uDiag : UDINT;  // 诊断字，16#0001_0152=tPT 负值已钳 0，0=无诊断事件 / Diag word, 16#0001_0152=negative tPT clamped to 0, 0=no diag event
END_VAR
VAR
    fbTon    : TON;   // 内建接通延时实例，承担单段计时内核 / Built-in TON instance, owns the per-segment timing kernel
    tPTClamp : TIME;  // 钳位后的预置总延时 [ms]，喂给内建实例 / Clamped preset total delay [ms], fed to the built-in instance
    tAccum   : TIME;  // 保持量累计 [ms]，跨暂停段保持 / Retained accumulation [ms], kept across pause segments
    tETLast  : TIME;  // 上一扫描周期的实时计时快照 [ms]，供断开拍冻结 / Last-scan elapsed snapshot [ms], frozen on the drop scan
    bRunPrev : BOOL;  // 上一扫描周期 bIN 快照，用于下降沿识别 / Previous-scan bIN snapshot, for falling-edge detection
    bDone    : BOOL;  // 累计到达内部锁存位 / Internal done latch
    xInit    : BOOL;  // 首扫初始化标志，FALSE=尚未完成上电初始化 / First-scan init flag, FALSE = power-on init not yet done
END_VAR

(*------------------------------------------------------------------------------
 * 段 1｜首扫初始化（历史教训④口径）：置于逻辑最前，首扫不产假 bQ
 *      First-scan init (lesson 4): placed at the very front, no false bQ on first scan
 *-----------------------------------------------------------------------------*)
IF NOT xInit THEN
    xInit    := TRUE;    // 置初始化完成标志 / Mark init as done
    tPTClamp := T#0s;    // 首扫钳位值归零，避免未初始化喂入 / Zero the clamp value on first scan
    tAccum   := T#0s;    // 首扫保持量清零 / Zero retained accumulation on first scan
    tETLast  := T#0s;    // 首扫计时快照清零 / Zero elapsed snapshot on first scan
    bRunPrev := FALSE;   // 首扫使能快照为 FALSE，杜绝假下降沿 / FALSE on first scan, no false falling edge
    bDone    := FALSE;   // 首扫到时位清零 / Clear done latch on first scan
    uDiag    := 16#0000_0000;  // 首扫诊断字清零 / Clear diag word on first scan
END_IF

(*------------------------------------------------------------------------------
 * 段 2｜PT 域校验与钳位：负 TIME 统一钳 0 并置信息码
 *      PT domain check and clamp: negative TIME unified to 0 with informational code
 *-----------------------------------------------------------------------------*)
IF tPT < T#0s THEN
    tPTClamp := T#0s;        // 负值钳位为 0 [ms] / Clamp negative to 0 [ms]
    uDiag    := 16#0001_0152;  // 信息码：PT 负值已钳 0 / Informational: negative PT clamped to 0
ELSE
    tPTClamp := tPT;         // 域内直通 / In-domain pass-through
    uDiag    := 16#0000_0000;  // 无诊断事件，清码 / No diag event, clear code
END_IF

(*------------------------------------------------------------------------------
 * 段 3｜复位类写入（前置，历史教训⑦）：bRESET 电平优先级最高，清零累计与
 *      到时位；即使同拍 bIN=TRUE 也走复位语义（段 5 内建实例随后重新起计时）
 *      Reset-class writes (front, lesson 7): level reset has top priority;
 *      even with bIN TRUE on the same scan, reset semantics wins
 *-----------------------------------------------------------------------------*)
IF bRESET THEN
    tAccum := T#0s;    // 清零保持量累计 [ms] / Clear retained accumulation [ms]
    bDone  := FALSE;   // 清零到时锁存位 / Clear done latch
END_IF

(*------------------------------------------------------------------------------
 * 段 4｜下降沿冻结（置位类，须在内建 TON 调用之前）：bIN 断开当拍，内建 TON
 *      将被本次调用清零，故取上一拍快照 tETLast 冻结累入保持量；
 *      复位拍与到时态不冻结（复位已清零、到时无未结段落）
 *      Falling-edge freeze (set-class, before the built-in TON call): on the
 *      scan bIN drops, the built-in TON will be zeroed by this very call, so
 *      the last-scan snapshot tETLast is frozen into the retention
 *-----------------------------------------------------------------------------*)
IF bRunPrev AND (NOT bIN) AND (NOT bDone) AND (NOT bRESET) THEN
    tAccum := tAccum + tETLast;  // 冻结上一拍实时计时入保持量 [ms] / Freeze last-scan elapsed into retention [ms]
END_IF

(*------------------------------------------------------------------------------
 * 段 5｜无条件刷新区（红线 R7）：TON 实例严禁进入任何 IF / CASE 分支；
 *      IN = 使能且未到时——到时后自动摘除使能，杜绝重复计时
 *      Unconditional refresh zone (red line R7): no instance call inside IF / CASE;
 *      IN = enabled AND not done, auto-detached after completion
 *-----------------------------------------------------------------------------*)
fbTon(IN := bIN AND (NOT bDone), PT := tPTClamp);  // 每扫描周期无条件喂入 / Feed unconditionally every scan

(*------------------------------------------------------------------------------
 * 段 6｜到时锁存（实例调用之后置位类写入，R24 教训）：完成拍把本段满程计时
 *      （此时 ET=钳位后 PT）累入保持量并锁存到时位
 *      Done latch (set-class write after the instance call, R24 lesson): on the
 *      completion scan, the full segment (ET = clamped PT) is frozen and done latched
 *-----------------------------------------------------------------------------*)
IF fbTon.Q AND (NOT bDone) THEN
    bDone  := TRUE;              // 锁存累计到达 / Latch accumulated-done
    tAccum := tAccum + fbTon.ET; // 本段满程计时累入保持量 [ms]（完成拍 ET=钳位后 PT）/ Full segment frozen into retention [ms], ET equals clamped PT on the completion scan
END_IF

(*------------------------------------------------------------------------------
 * 段 7｜输出组合：运行中 = 保持量 + 本段实时值；暂停/到时/复位 = 仅保持量
 *      Output composition: running = retention + live segment; else retention only
 *-----------------------------------------------------------------------------*)
IF bIN AND (NOT bDone) THEN
    tET := tAccum + fbTon.ET;  // 运行中输出 [ms] / Live output while running [ms]
ELSE
    tET := tAccum;             // 暂停/到时/复位输出仅保持量 [ms] / Paused/done/reset output, retention only [ms]
END_IF
bQ := bDone;                 // 累计到达输出 / Accumulated-done output

(*------------------------------------------------------------------------------
 * 段 8｜周期快照落盘：本拍使能与实时计时供下一拍下降沿冻结取用
 *      Per-scan snapshot: this scan's enable and live elapsed feed next scan's freeze
 *-----------------------------------------------------------------------------*)
bRunPrev := bIN;      // 快照本拍使能 / Snapshot this scan's enable
tETLast  := fbTon.ET; // 快照本拍实时计时 [ms] / Snapshot this scan's live elapsed [ms]
END_FUNCTION_BLOCK

(* ---- FB_DL_RTrigEx.st ---- *)
(*==============================================================================
 * 组件名称 (Component)  : FB_DL_RTrigEx
 * 所属子库 (Sublibrary) : DL_Base
 * 当前版本 (Version)    : 1.0.0
 * 兼容性   (Platform)   : CODESYS 3.5 / TwinCAT 3 / 汇川 InoProShop / Machine Expert
 *                         仅依赖 Standard.library（R_TRIG），零厂商方言
 * 功能描述 (Function)   : 上升沿检测防御包装。内部委托 IEC 61131-3 标准 R_TRIG
 *                         实例完成沿检测内核，外围统一首扫时序行为（首扫按 CLK
 *                         当前值建立基线、不产假边沿）并保证输出严格单拍。
 * 溯源     (Origin)     : IEC 61131-3 标准语义的道莅防御性实现
 *                         （接口语义由 IEC 61131-3 定义，clean-room 重写，
 *                         参考公开标准条款）
 * 码位     (Diag Codes) : 无错误码（纯语义包装，输入为单布尔量，无域可校验）
 *                         本件不占用 014D~015D / 0226~022B 任何码位
 * 类型裁定 (Type Note)  : 本件无诊断字引脚，错误码声明以本节替代
 * 依赖     (Depends)    : 无 DL_ 内部依赖；Standard.library: R_TRIG
 * 红线自检 (Redline)    : R1 ✓ 零全局变量与外部变量引用 ｜ R2 ✓ 零物理 IO 地址直写
 *                         R3 ✓ 纯 IEC 61131-3 ｜ R4 ✓ 首扫不假触发+单拍输出
 *                         R5 ✓ 全变量中英双语同行注释 ｜ R6 N/A（无顺序状态机，见下）
 *                         R7 ✓ R_TRIG 实例主体无条件周期刷新
 * 说明     (Note)       : R6 标注 N/A —— 本组件为单步沿检测，不存在顺序状态机，
 *                         无 CASE 可写；非法状态不可能出现（唯一状态即"运行"），
 *                         故以本节说明替代 ELSE 兜底，符合"无状态机则标注 N/A"口径。
 * 防御行为声明 (Defense): ① 首扫不产假边沿：部分平台 R_TRIG 首扫在 CLK=TRUE 时会
 *                           输出 Q=TRUE（平台行为不一致），本件统一为首扫抑制一拍，
 *                           从第二拍起交付标准沿语义；
 *                         ② 单拍输出保证：bQ 仅在真实上升沿所在扫描周期为 TRUE，
 *                           下一拍自动归 FALSE（由内建 R_TRIG 语义保证）；
 *                         ③ 上电即处于 TRUE 的 CLK 不算沿（与"沿=跳变"定义一致）。
 * 修订历史 (Revision)   :
 *   2026-11-16  v1.0.0  首版入库（R14 批 1 · T0 快车道）
 *============================================================================*)
FUNCTION_BLOCK FB_DL_RTrigEx
VAR_INPUT
    bCLK : BOOL;  // 时钟输入，检测其低→高跳变 / Clock input, detects its low-to-high transition
END_VAR
VAR_OUTPUT
    bQ : BOOL;    // 单拍上升沿脉冲，仅在跳变所在扫描周期为 TRUE / One-scan rising-edge pulse, TRUE only on the scan of the transition
END_VAR
VAR
    fbTrig : R_TRIG;  // 内建上升沿检测实例，承担沿检测内核 / Built-in rising-edge instance, owns the edge-detection kernel
    xInit  : BOOL;    // 首扫初始化标志，FALSE=尚未完成上电初始化 / First-scan init flag, FALSE = power-on init not yet done
END_VAR

(*------------------------------------------------------------------------------
 * 段 1｜无条件刷新区（红线 R7）：R_TRIG 实例严禁进入任何 IF / CASE 分支
 *      Unconditional refresh zone (red line R7): no instance call inside IF / CASE
 *-----------------------------------------------------------------------------*)
fbTrig(CLK := bCLK);  // 每扫描周期无条件喂入时钟 / Feed clock unconditionally every scan

(*------------------------------------------------------------------------------
 * 段 2｜首扫初始化（历史教训⑤口径）：置于逻辑最前，首扫抑制内建实例输出一拍，
 *      统一各平台 R_TRIG 首扫行为差异
 *      First-scan init (lesson 5): placed at the very front; suppress the built-in
 *      output for one scan to unify cross-platform first-scan behavior
 *-----------------------------------------------------------------------------*)
IF NOT xInit THEN
    xInit := TRUE;   // 置初始化完成标志 / Mark init as done
    bQ    := FALSE;  // 首扫强制 FALSE，不产假边沿 / Force FALSE on first scan, no false edge
ELSE
    bQ := fbTrig.Q;  // 非首扫：直通内建沿检测输出（天然单拍）/ Non-first scan: pass through built-in edge output (single-scan by nature)
END_IF
END_FUNCTION_BLOCK

(* ---- FB_DL_RuntimeMeter.st ---- *)
(*==============================================================================
 * 组件名称 (Component)  : FB_DL_RuntimeMeter
 * 所属子库 (Sublibrary) : DL_Base
 * 当前版本 (Version)    : 1.0.0
 * 兼容性   (Platform)   : CODESYS 3.5 / TwinCAT 3 / 汇川 InoProShop / Machine Expert
 *                         仅依赖 Standard.library（R_TRIG），零平台时刻函数
 * 功能描述 (Function)   : 设备累计运行时间（分钟 / 小时双口径）与启动次数统计，
 *                         带保养间隔到期预警。时间增量由调用方注入，本块零平台依赖。
 *                         采用"秒 + 毫秒进位缓存"的整数化累加，不做逐周期浮点累加，
 *                         从根上消除浮点漂移（与滑动平均的整数化思想同源）。
 *                         保养到期锁存至确认沿；启动计数达上限饱和停增不回绕。
 * 开源溯源 (Origin)     : 原创实现。运行小时表 + 保养计数的功能组合为工业界通行做法，
 *                         整数化累加与注入式时间设计为本库既有范式，未复制任何源码。
 * 本文件内含       : FB    FB_DL_RuntimeMeter（单 POU，无配套类型）
 * 依赖     (Depends)    : 无 DL_ 内部依赖；Standard.library: R_TRIG
 * 红线自检 (Redline)    : R1 ✓ 禁用全局存储与物理寻址 ｜ R2 ✓ 无地址直写
 *                         R3 ✓ 纯 IEC 61131-3，零平台时刻函数 ｜ R4 ✓ 增量拒收 + 乘法溢出钳位 + 结构性除零论证
 *                         R5 ✓ 全变量中英双语同行注释 ｜ R6 N/A（纯累计统计，无状态转移）
 *                         R7 ✓ 三 R_TRIG 主体最前部无条件刷新 ｜ R8 ✓ 换算系数全部常量化
 *
 * 【断电保持提示 / Retain hint（边界 B9）】
 *   本块全部累计量若不声明为断电保持类型，重新上电即归零，保养预警与启动次数随之丢失。
 *   推荐调用方把本 FB 的实例声明为断电保持变量。
 *   All accumulators are lost on power cycle unless the caller declares the instance retentive.
 *
 * 【除零结构性豁免 / Structural divide-by-zero exemption（边界 B7）】
 *   fRunHours 的除数为常量 3600 秒/小时，编译期恒大于零，不存在运行期为零的可能，
 *   故不设前置判断；uMaintRemainMin 的除数为常量 60 秒/分钟，同理。
 *   The divisors are compile-time positive constants, so no runtime guard is required.
 *
 * 修订历史 (Revision)   :
 *   2026-11-14  v1.0.0  首版入库（Phase 1 第二轮 · Level 0 批次 A）
 *============================================================================*)
FUNCTION_BLOCK FB_DL_RuntimeMeter
VAR_INPUT
    bRunning          : BOOL;                  // 设备运行反馈（电平，TRUE 期间累计时间）/ Equipment running feedback, level
    uDeltaTimeMs      : UDINT;                 // 本任务周期耗时 [ms]，调用方注入 / Cycle time in ms, caller-provided
    uMaintIntervalMin : UDINT := UDINT#0;      // 保养间隔 [min]，0 = 关闭保养预警 / Maintenance interval [min], 0 = disabled
    bMaintAck         : BOOL;                  // 上升沿：保养确认，重置保养计时 / Rising edge: acknowledge maintenance
    bReset            : BOOL;                  // 上升沿：清零全部累计 / Rising edge: clear all totals
END_VAR
VAR_OUTPUT
    uRunTotalMin     : UDINT;   // 累计运行时间 [min] / Total runtime in minutes
    fRunHours        : REAL;    // 累计运行小时 [h]（HMI 直显口径）/ Total runtime in hours for HMI
    nStartCount      : UDINT;   // 累计启动次数 [次] / Accumulated start count [count]
    bMaintDue        : BOOL;    // 保养到期（锁存至确认）/ Maintenance due, latched until acknowledged
    uMaintRemainMin  : UDINT;   // 距下次保养剩余 [min]，未启用时为 0 / Minutes to next maintenance, 0 when disabled
    uErrorId         : UDINT;   // 故障码，0 = 无故障 / Error code, 0 = no error
END_VAR
VAR
    uTotalSec        : UDINT;   // 累计运行秒 [s] / Total runtime seconds [s]
    uSinceMaintSec   : UDINT;   // 距上次保养累计秒 [s] / Seconds since last maintenance [s]
    uMsCarry         : UDINT;   // 毫秒进位缓存 [ms] / Millisecond carry buffer [ms]
    fbTrigRun        : R_TRIG;  // 启动上升沿检测实例 / Start rising edge detector instance
    fbTrigMaintAck   : R_TRIG;  // 保养确认上升沿检测实例 / Maintenance ack rising edge detector instance
    fbTrigReset      : R_TRIG;  // 复位上升沿检测实例 / Reset rising edge detector instance
    uMaintIntEff     : UDINT;   // 钳位后的保养间隔 [min] / Clamped maintenance interval [min]
    uMaintThreshSec  : UDINT;   // 保养到期门槛秒数 [s] / Maintenance due threshold in seconds
    uCarrySec        : UDINT;   // 本周期可折算的整秒数 [s] / Whole seconds derivable this cycle
END_VAR
VAR CONSTANT
    DL_RT_SEC_PER_MIN   : UDINT := 60;             // 每分钟秒数 [s/min] / Seconds per minute
    DL_RT_SEC_PER_HOUR  : UDINT := 3600;           // 每小时秒数 [s/h] / Seconds per hour
    DL_RT_MS_PER_SEC    : UDINT := 1000;           // 每秒毫秒数 [ms/s] / Milliseconds per second
    DL_RT_COUNT_MAX     : UDINT := 16#FFFF_FFFE;   // 启动计数饱和上限 [次] / Start count saturation limit
    DL_RT_DELTA_MAX     : UDINT := 3600000;        // 单周期合理上限 [ms] / Sanity cap per cycle [ms]
    DL_RT_MAINT_INT_MAX : UDINT := 525600;         // 保养间隔上限 [min]，一年，防乘法溢出 / Interval cap [min], one year
END_VAR

(*------------------------------------------------------------------------------
 * 段 1｜无条件刷新区（红线 R7）：三个边沿实例位于主体最前部，严禁进入 IF / CASE
 *      Unconditional refresh zone: all three edge instances run at the very top
 *-----------------------------------------------------------------------------*)
fbTrigRun(CLK := bRunning);
fbTrigMaintAck(CLK := bMaintAck);
fbTrigReset(CLK := bReset);

(*------------------------------------------------------------------------------
 * 段 2｜故障码本周期清零：错误码只描述当前周期事实
 *      Error code is cleared every scan: it reports the current cycle only
 *-----------------------------------------------------------------------------*)
uErrorId := 16#0000_0000;

(*------------------------------------------------------------------------------
 * 段 3｜复位语义（边界 B8）：全部累计归零，故障码同时清除，口径统一
 *      Reset: every total goes to zero together with the error code
 *-----------------------------------------------------------------------------*)
IF fbTrigReset.Q THEN
    uTotalSec       := UDINT#0;
    uSinceMaintSec  := UDINT#0;
    uMsCarry        := UDINT#0;
    uRunTotalMin    := UDINT#0;
    fRunHours       := 0.0;
    nStartCount     := UDINT#0;
    bMaintDue       := FALSE;
    uMaintRemainMin := UDINT#0;
END_IF

(*------------------------------------------------------------------------------
 * 段 4｜保养间隔钳位（边界 B6）：上限一年，防止分钟折算秒时乘法溢出
 *      Interval clamping: one year cap prevents overflow in the minute-to-second product
 *-----------------------------------------------------------------------------*)
IF uMaintIntervalMin > DL_RT_MAINT_INT_MAX THEN
    uMaintIntEff := DL_RT_MAINT_INT_MAX;
    uErrorId     := 16#0001_0001;
ELSE
    uMaintIntEff := uMaintIntervalMin;
END_IF

uMaintThreshSec := uMaintIntEff * DL_RT_SEC_PER_MIN;

(*------------------------------------------------------------------------------
 * 段 5｜增量防御（边界 B3）：零增量与超上限增量均不计入，口径与周期测量块一致
 *      Delta defence: zero and over-limit deltas are ignored, same policy as the cycle block
 *-----------------------------------------------------------------------------*)
IF (uDeltaTimeMs > UDINT#0) AND (uDeltaTimeMs <= DL_RT_DELTA_MAX) THEN

    IF bRunning THEN
        (*----------------------------------------------------------------------
         * 段 6｜毫秒进位累加（边界 B2）：先把毫秒攒够整秒，再折算进秒计数
         *      Millisecond carry: accumulate to whole seconds before folding into the counters
         *      避免每周期浮点累加，长期运行不产生漂移；进位缓存保留不足一秒的余量
         *      No per-cycle float accumulation, so no long-term drift is possible
         *---------------------------------------------------------------------*)
        uMsCarry := uMsCarry + uDeltaTimeMs;

        IF uMsCarry >= DL_RT_MS_PER_SEC THEN
            (* 除数 1000 为编译期正的常量，结构性免除零判断（见头注释） *)
            (* The divisor 1000 is a compile-time positive constant, structurally safe *)
            uCarrySec  := uMsCarry / DL_RT_MS_PER_SEC;
            uMsCarry   := uMsCarry - (uCarrySec * DL_RT_MS_PER_SEC);
            uTotalSec  := uTotalSec + uCarrySec;
            uSinceMaintSec := uSinceMaintSec + uCarrySec;
        END_IF
    END_IF

ELSE
    uErrorId := 16#0001_0008;
END_IF

(*------------------------------------------------------------------------------
 * 段 7｜启动计数（边界 B4）：上升沿计数，达上限饱和停增，绝不回绕
 *      Start count: rising edge increments, saturation instead of wrap-around
 *-----------------------------------------------------------------------------*)
IF fbTrigRun.Q THEN
    IF nStartCount < DL_RT_COUNT_MAX THEN
        nStartCount := nStartCount + UDINT#1;
    ELSE
        uErrorId := 16#0001_0007;
    END_IF
END_IF

(*------------------------------------------------------------------------------
 * 段 8｜保养预警（边界 B5）：到期锁存，确认沿清零计时并解除锁存
 *      Maintenance warning: latched on due, cleared by the acknowledge edge
 *-----------------------------------------------------------------------------*)
IF uMaintIntEff = UDINT#0 THEN
    (* 功能关闭：不预警、不显示剩余，历史保养计时保留不影响累计口径 *)
    (* Function disabled: no warning, no remaining display, history is kept *)
    bMaintDue       := FALSE;
    uMaintRemainMin := UDINT#0;
ELSE
    IF uSinceMaintSec >= uMaintThreshSec THEN
        bMaintDue := TRUE;
    END_IF

    IF fbTrigMaintAck.Q THEN
        bMaintDue      := FALSE;
        uSinceMaintSec := UDINT#0;
    END_IF

    IF uSinceMaintSec >= uMaintThreshSec THEN
        uMaintRemainMin := UDINT#0;
    ELSE
        (* 除数 60 为编译期正的常量，结构性免除零判断（见头注释） *)
        (* The divisor 60 is a compile-time positive constant, structurally safe *)
        uMaintRemainMin := (uMaintThreshSec - uSinceMaintSec) / DL_RT_SEC_PER_MIN;
    END_IF
END_IF

(*------------------------------------------------------------------------------
 * 段 9｜输出刷新：分钟取整下取整口径，小时保留小数供 HMI 直显
 *      Output refresh: minutes are truncated, hours keep the fractional part for HMI
 *      除数 3600 为编译期正的常量，结构性免除零判断（边界 B7）
 *      The divisor 3600 is a compile-time positive constant, structurally safe
 *-----------------------------------------------------------------------------*)
uRunTotalMin := uTotalSec / DL_RT_SEC_PER_MIN;
fRunHours    := UDINT_TO_REAL(uTotalSec) / UDINT_TO_REAL(DL_RT_SEC_PER_HOUR);
END_FUNCTION_BLOCK

(* ---- FB_DL_SamplingTrigger.st ---- *)
(*
    组件名称 : FB_DL_SamplingTrigger
    所属子库 : DL_Base
    当前版本 : 1.0.0
    兼 容 性 : CODESYS V3.5+ / TwinCAT 3 / 汇川 InoProShop；仅依赖 Standard.library
    功能描述 : 均匀采样节拍源，输出单拍采样沿 + 样本序号 + 理论/实际时基账目 + 漂移告警，供趋势记录使用。
              取舍 ①：理论时长用「样本序号 × 周期」重算，而不是每拍累加周期 —— 累加式在每一次「定时器命中
              晚一个扫描周期」时都会永久吞掉那点误差，跑一天能差出几十毫秒；序号重算则误差不累积，
              这正是「无漂移」三个字的来源。
              取舍 ②：扫描周期增量由调用方注入（tDelta），不调平台时刻函数 —— 与库内 CycleTimeMeasure 同一纪律，
              换平台不必改代码，也让副程序内的假节拍可复现测试。
              取舍 ③：tDelta ≤ 0 时本拍不累加实际时基 —— 首扫或注入错误时，凭空加一个增量会让 tActual
              从第一拍就偏；本件宁可少记一拍，也不伪造时间。
              取舍 ④：漂移只提示不重置 —— 重置会让「真实时基丢失」这个事实消失在账目里；留着偏差，
              上位机每次取数都能看到它。
              取舍 ⑤：与 FB_DL_PulseGenerator 的边界 —— 那件出占空比可调的方波；本件只出采样沿与时基账目。
    开源溯源 : 原创实现（T0-2 变体线）。无外部源码参考，码位、漂移阈值、回绕策略 100% 自有。；本件为 IEC 61131-3 标准语义的道莅防御性实现（原创实现，零外部源码复制）。
    本文件内含 : FUNCTION_BLOCK FB_DL_SamplingTrigger（单 POU，无配套类型）
    依 赖 : 无 DL_ 内部依赖；Standard.library: TON / R_TRIG
    红线自检 : R1 ✓ 零全局变量与外部变量 ｜ R2 ✓ 零物理 IO 地址
              R3 ✓ 纯 IEC 61131-3 ｜ R4 ✓ 周期闸 + 增量闸 + 序号回绕 + 理论值溢出预判 + 漂移双侧直比
              R5 ✓ 全变量中英双语同行注释 ｜ R6 N/A 无顺序状态机（纯节拍累加），头注释已写明理由
              R7 ✓ TON / R_TRIG 实例在主体最前部无条件刷新，IN 含使能与复位，保证重新使能不产生假沿
              R8 ✓ 周期下限、增量上限、漂移阈值全常量化
    错误码   : 16#0001_0456 [信息级] 累计漂移超阈值，只提示不重置，bError = FALSE
               16#0001_0457 [信息级] 样本序号回绕归零，bError = FALSE
               16#0001_039F [故障级] 采样周期非法已钳至 1ms 继续，bError = TRUE
               16#0001_03A0 [故障级] 扫描周期增量非法（≤ 0 或超上限），本拍不计入实际时基，bError = TRUE
               16#0001_03A1 [故障级] 预留禁用（不得挪用）
    码位总账 : 16#0001_0456 用 / 16#0001_0457 用 ｜ 16#0001_039F 用 / 16#0001_03A0 用 / 16#0001_03A1 预留
    遗留假设 : ① TIME 为 32 位有符号毫秒口径；tActual 的加法已做溢出预判（R54：比较式内不出现加乘），
              超上限时保持上拍值不累加，故无回绕路径。该口径未在 InoProShop 实测。
              ② 漂移判据在 DINT 毫秒域做双侧直比（nDiff > +阈 OR nDiff < −阈），不用 ABS 单侧，
              避免差值在极端情形下取绝对值回绕（有符号整数边界纪律）。
    修订历史 :
        2026-11-16  v1.0.0  首版，R21 批次 4 入库
*)
FUNCTION_BLOCK FB_DL_SamplingTrigger
VAR_INPUT
    bEnable         : BOOL := TRUE;      // 使能，FALSE 时不产生样本但定时器仍刷新 / enable, FALSE stops the samples while the timer keeps refreshing
    tInterval       : TIME := T#1S;      // 采样周期，≤ 0 时钳至 1ms [ms] / sampling period, clamped to one millisecond [ms]
    tDelta          : TIME;              // 调用方注入的扫描周期增量，必须 > 0 [ms] / scan time increment injected by the caller, must be positive [ms]
    bReset          : BOOL;              // 上升沿清序号与时基账目 / rising edge clears the sample number and the time accounts
END_VAR
VAR_OUTPUT
    bSample         : BOOL;              // 单拍采样沿，仅 TRUE 一个扫描周期 / single scan sample edge
    uSampleNo       : UDINT;             // 样本序号，1 起；回绕时归零 [个] / sample number starting at one, wrapped to zero on overflow [count]
    tTheoretical    : TIME;              // 理论累计时长 = 序号 × 周期 [ms] / theoretical elapsed time, samples times the period [ms]
    tActual         : TIME;              // 注入增量累计的实际时长 [ms] / actual elapsed time accumulated from the injected increments [ms]
    bDrift          : BOOL;              // 偏差超阈值，锁存至复位 / TRUE when the deviation exceeds the threshold, latched until reset
    eErr            : UDINT;             // 错误码，0=正常；16#0001_04XX 信息级 / 16#0001_03XX 故障级 / error id, 0=ok
    bError          : BOOL;              // 故障级标志 / fault flag
END_VAR
VAR
    fbTimer         : TON;               // 采样周期定时器，主体最前部无条件刷新 / sampling timer, refreshed unconditionally at the top
    rtSample        : R_TRIG;            // 定时器完成位上升沿，主体最前部无条件刷新 / rising edge of the timer output, refreshed unconditionally
    tIntervalEff    : TIME;              // 钳位后的采样周期 [ms] / clamped sampling period [ms]
    bTimerIn        : BOOL;              // 定时器输入，含使能与复位 / timer input including the enable and the reset
    bDeltaOk        : BOOL;              // 本拍增量是否可用于累加 / whether the increment may be accumulated this scan
    nIntervalMs     : DINT;              // 采样周期的毫秒值 [ms] / sampling period in milliseconds [ms]
    nDeltaMs        : DINT;              // 增量的毫秒值 [ms] / increment in milliseconds [ms]
    nActualMs       : DINT;              // 实际时基的毫秒值 [ms] / actual elapsed time in milliseconds [ms]
    nDiffMs         : DINT;              // 实际与理论的毫秒偏差，可正可负 [ms] / deviation between the actual and the theoretical time, signed [ms]
    nMaxSamples     : DINT;              // 理论值不溢出的最大样本数 [个] / largest sample number whose product stays in range [count]
END_VAR
VAR CONSTANT
    DL_SAMPLE_INT_MIN   : TIME := T#1MS;                  // 采样周期下限 [ms] / sampling period lower bound [ms]
    DL_SAMPLE_DRIFT_MAX : TIME := T#200MS;                // 漂移告警阈值 [ms] / drift warning threshold [ms]
    DL_DELTA_MAX        : TIME := T#10S;                  // 增量上限，超此值视为任务卡顿 [ms] / increment upper bound, beyond it the task stalled [ms]
    DL_TIME_ZERO        : TIME := T#0S;                   // 零时长哨兵 [ms] / zero duration sentinel [ms]
    DL_TIME_MS_MAX      : DINT := 2147483647;             // TIME 毫秒上限，加法预判用 [ms] / TIME millisecond bound used by the addition prediction [ms]
    DL_DINT_ZERO        : DINT := 0;                      // 整数零哨兵 [无量纲] / integer zero sentinel [dimensionless]
    DL_UDINT_MAX        : UDINT := 16#FFFF_FFFF;          // 序号上限 [个] / sample number upper bound [count]
    DL_UDINT_ZERO       : UDINT := 0;                     // 序号零哨兵 [个] / sample number zero sentinel [count]
    DL_ERR_NONE         : UDINT := 16#0000_0000;          // 无故障 / no error
END_VAR

// 段 0｜错误状态预置与单拍标志清销 / segment 0, preset the error state and clear the single scan flag
eErr    := DL_ERR_NONE;                      // 预置无错误 / preset no error
bError  := FALSE;                            // 预置无故障 / preset no fault
bSample := FALSE;                            // 单拍标志每拍先销，防「只置不销」/ the single scan flag is cleared first, never left latched

// 段 1｜采样周期闸：非法则钳 1ms 继续，不停机 / segment 1, period gate, clamp instead of stopping
IF tInterval <= DL_TIME_ZERO THEN
    tIntervalEff := DL_SAMPLE_INT_MIN;       // 钳到最小周期 / clamp to the smallest period
    eErr   := 16#0001_039F;                  // 采样周期非法已钳位（故障级）/ illegal period clamped, fault level
    bError := TRUE;                          // 置故障标志 / raise the fault flag
ELSE
    tIntervalEff := tInterval;               // 正常值 / a healthy value
END_IF

// 段 2｜定时器与边沿无条件刷新：IN 含使能与复位，重新使能时不会留下假沿 / segment 2, unconditional refresh
bTimerIn := bEnable AND NOT bReset;
fbTimer ( IN := bTimerIn, PT := tIntervalEff );
rtSample( CLK := fbTimer.Q );

// 段 3｜增量闸：≤ 0 视为首扫或注入错误，本拍不累加也不出样本 / segment 3, increment gate
bDeltaOk := tDelta > DL_TIME_ZERO;
IF NOT bDeltaOk THEN
    eErr   := 16#0001_03A0;                  // 周期增量非法（故障级）/ illegal increment, fault level
    bError := TRUE;                          // 置故障标志 / raise the fault flag
ELSIF tDelta > DL_DELTA_MAX THEN
    bDrift := TRUE;                          // 任务卡顿，累加但置漂移 / the task stalled, accumulate and flag the drift
    eErr   := 16#0001_03A0;                  // 同一判据同一码（增量不可信）/ the same cause shares one code
    bError := TRUE;                          // 置故障标志 / raise the fault flag
END_IF

// 段 4｜复位沿：清序号与时基账目 / segment 4, reset clears the counter and both time accounts
IF bReset THEN
    uSampleNo    := DL_UDINT_ZERO;           // 序号归零 / clear the sample number
    tActual      := DL_TIME_ZERO;            // 实际时基归零 / clear the actual time
    tTheoretical := DL_TIME_ZERO;            // 理论时基归零 / clear the theoretical time
    bDrift       := FALSE;                   // 解除漂移锁存 / release the drift latch
END_IF

// 段 5｜采样沿与序号推进 / segment 5, sample edge and number advance
IF rtSample.Q AND bEnable THEN
    bSample := TRUE;                         // 单拍采样沿 / the single scan sample edge
    IF uSampleNo >= DL_UDINT_MAX THEN
        uSampleNo := DL_UDINT_ZERO;          // 回绕归零，理论值随之重算 / wrap to zero, the theoretical time restarts with it
        IF eErr = DL_ERR_NONE THEN
            eErr := 16#0001_0457;            // 样本序号回绕（信息级）/ sample number wrapped, info level
        END_IF
    ELSE
        uSampleNo := uSampleNo + 1;          // 序号自增，首样本为 1 / advance, the first sample is one
    END_IF
END_IF

// 段 6｜实际时基累加：先做溢出预判，比较式内不出现加乘（R54）/ segment 6, actual time accumulation with an overflow prediction
IF bDeltaOk THEN
    nActualMs := TIME_TO_DINT(tActual);      // 当前实际时基 [ms] / current actual time [ms]
    nDeltaMs  := TIME_TO_DINT(tDelta);       // 本拍增量 [ms] / the increment of this scan [ms]
    IF nActualMs > DL_TIME_MS_MAX - nDeltaMs THEN
        tActual := DINT_TO_TIME(DL_TIME_MS_MAX);   // 顶到上限，保持可观测而不回绕 / cap at the bound instead of wrapping
    ELSE
        tActual := DINT_TO_TIME(nActualMs + nDeltaMs);   // 正常累加 / normal accumulation
    END_IF
END_IF

// 段 7｜理论时基：序号 × 周期重算，误差不累积；先算可容纳样本数防溢出 / segment 7, theoretical time recomputed from the number
nIntervalMs := TIME_TO_DINT(tIntervalEff);   // 周期毫秒值，闸后恒 ≥ 1 / the period is at least one millisecond after the gate
IF nIntervalMs > DL_DINT_ZERO THEN
    nMaxSamples := DL_TIME_MS_MAX / nIntervalMs;   // 不溢出的最大样本数 / the largest number that keeps the product in range
    IF uSampleNo <= DINT_TO_UDINT(nMaxSamples) THEN
        tTheoretical := DINT_TO_TIME(nIntervalMs * UDINT_TO_DINT(uSampleNo));   // 理论值 = 序号 × 周期 / theoretical equals the number times the period
    END_IF
END_IF

// 段 8｜漂移判据：DINT 毫秒域双侧直比，禁 ABS 单侧 / segment 8, drift test with a two sided comparison
nDiffMs := TIME_TO_DINT(tActual) - TIME_TO_DINT(tTheoretical);
IF (nDiffMs > TIME_TO_DINT(DL_SAMPLE_DRIFT_MAX)) OR (nDiffMs < (DL_DINT_ZERO - TIME_TO_DINT(DL_SAMPLE_DRIFT_MAX))) THEN
    bDrift := TRUE;                          // 漂移锁存，不重置（重置会掩盖时基丢失）/ latch the drift, a reset would hide the lost time base
    IF eErr = DL_ERR_NONE THEN
        eErr := 16#0001_0456;                // 累计漂移超阈值（信息级）/ accumulated drift, info level
    END_IF
END_IF
END_FUNCTION_BLOCK
